REGION Network 3: Convoyeur 02
   RUNG wire#powerrail
      #Convoyeur_Hippodrome_2(x_Marche_auto := wire#w1, x_Arret_auto := wire#w2, x_Defaut_externe := "Bits_Globaux".x_Defaut_bloquant, x_enService := "Bits_Globaux".x_En_service, x_Marche_manu := "Tch_HMI".Tch_Manu[50], x_Arret_Manu := "Tch_HMI".Tch_Manu[51], x_Retour_defaut_thermique := "I_Def_Thermique_CV02_hyppo", DB_Convoyeur_DATA := "DB_Convoyeurs_Hipp".Convoyeur[2], Defaut =>)
   END_RUNG
   RUNG wire#powerrail
      Contact( "Bits_Globaux".x_En_cycle_auto )
   END_RUNG wire#w1
   RUNG wire#powerrail
      Contact( "Bits_Globaux".x_Demo_Hippo_en_cours )
   END_RUNG wire#w1
   RUNG wire#powerrail
      Contact( "Tch_HMI".Tch_Acy )
   END_RUNG wire#w2
   RUNG wire#powerrail
      Contact( #x_All_stations_empty )
   END_RUNG wire#w2
   // the same network as SCL:
   #Convoyeur_Hippodrome_2(x_Defaut_externe := "Bits_Globaux".x_Defaut_bloquant,   // "Convoyeur_Hippodrome"
                           x_enService := "Bits_Globaux".x_En_service,
                           x_Marche_auto := "Bits_Globaux".x_En_cycle_auto OR "Bits_Globaux".x_Demo_Hippo_en_cours,
                           x_Marche_manu := "Tch_HMI".Tch_Manu[50],
                           x_Arret_auto := "Tch_HMI".Tch_Acy OR #x_All_stations_empty,
                           x_Arret_Manu := "Tch_HMI".Tch_Manu[51],
                           x_Retour_defaut_thermique := "I_Def_Thermique_CV02_hyppo",
                           DB_Convoyeur_DATA := "DB_Convoyeurs_Hipp".Convoyeur[2]);
END_REGION

REGION Network 4: Convoyeur 03
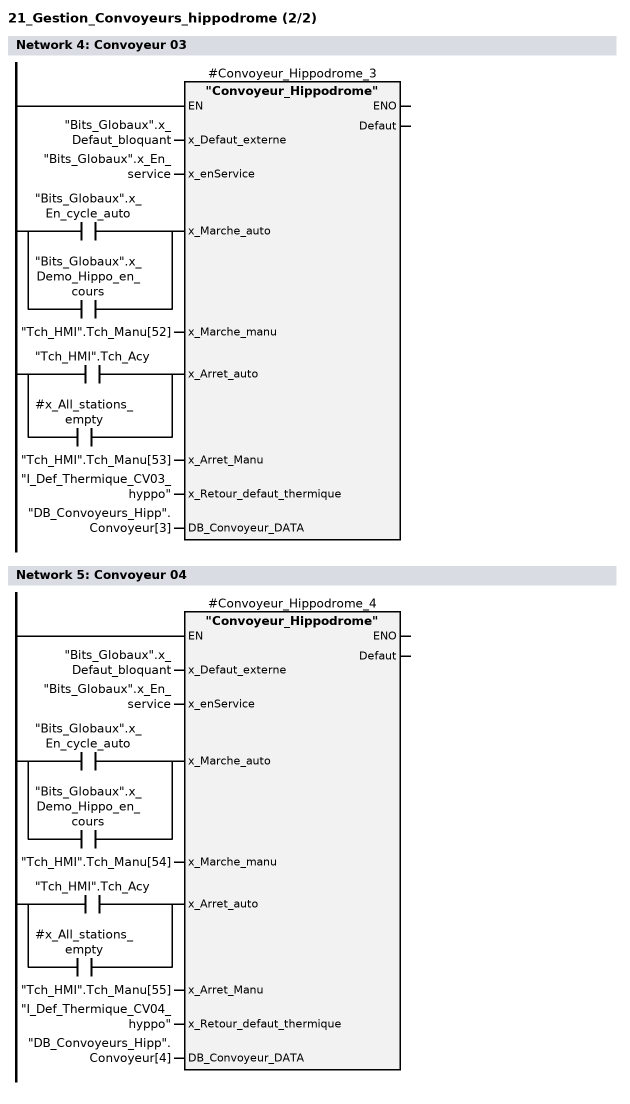
   RUNG wire#powerrail
      #Convoyeur_Hippodrome_3(x_Marche_auto := wire#w1, x_Arret_auto := wire#w2, x_Defaut_externe := "Bits_Globaux".x_Defaut_bloquant, x_enService := "Bits_Globaux".x_En_service, x_Marche_manu := "Tch_HMI".Tch_Manu[52], x_Arret_Manu := "Tch_HMI".Tch_Manu[53], x_Retour_defaut_thermique := "I_Def_Thermique_CV03_hyppo", DB_Convoyeur_DATA := "DB_Convoyeurs_Hipp".Convoyeur[3], Defaut =>)
   END_RUNG
   RUNG wire#powerrail
      Contact( "Bits_Globaux".x_En_cycle_auto )
   END_RUNG wire#w1
   RUNG wire#powerrail
      Contact( "Bits_Globaux".x_Demo_Hippo_en_cours )
   END_RUNG wire#w1
   RUNG wire#powerrail
      Contact( "Tch_HMI".Tch_Acy )
   END_RUNG wire#w2
   RUNG wire#powerrail
      Contact( #x_All_stations_empty )
   END_RUNG wire#w2
   // the same network as SCL:
   #Convoyeur_Hippodrome_3(x_Defaut_externe := "Bits_Globaux".x_Defaut_bloquant,   // "Convoyeur_Hippodrome"
                           x_enService := "Bits_Globaux".x_En_service,
                           x_Marche_auto := "Bits_Globaux".x_En_cycle_auto OR "Bits_Globaux".x_Demo_Hippo_en_cours,
                           x_Marche_manu := "Tch_HMI".Tch_Manu[52],
                           x_Arret_auto := "Tch_HMI".Tch_Acy OR #x_All_stations_empty,
                           x_Arret_Manu := "Tch_HMI".Tch_Manu[53],
                           x_Retour_defaut_thermique := "I_Def_Thermique_CV03_hyppo",
                           DB_Convoyeur_DATA := "DB_Convoyeurs_Hipp".Convoyeur[3]);
END_REGION

REGION Network 5: Convoyeur 04
   RUNG wire#powerrail
      #Convoyeur_Hippodrome_4(x_Marche_auto := wire#w1, x_Arret_auto := wire#w2, x_Defaut_externe := "Bits_Globaux".x_Defaut_bloquant, x_enService := "Bits_Globaux".x_En_service, x_Marche_manu := "Tch_HMI".Tch_Manu[54], x_Arret_Manu := "Tch_HMI".Tch_Manu[55], x_Retour_defaut_thermique := "I_Def_Thermique_CV04_hyppo", DB_Convoyeur_DATA := "DB_Convoyeurs_Hipp".Convoyeur[4], Defaut =>)
   END_RUNG
   RUNG wire#powerrail
      Contact( "Bits_Globaux".x_En_cycle_auto )
   END_RUNG wire#w1
   RUNG wire#powerrail
      Contact( "Bits_Globaux".x_Demo_Hippo_en_cours )
   END_RUNG wire#w1
   RUNG wire#powerrail
      Contact( "Tch_HMI".Tch_Acy )
   END_RUNG wire#w2
   RUNG wire#powerrail
      Contact( #x_All_stations_empty )
   END_RUNG wire#w2
   // the same network as SCL:
   #Convoyeur_Hippodrome_4(x_Defaut_externe := "Bits_Globaux".x_Defaut_bloquant,   // "Convoyeur_Hippodrome"
                           x_enService := "Bits_Globaux".x_En_service,
                           x_Marche_auto := "Bits_Globaux".x_En_cycle_auto OR "Bits_Globaux".x_Demo_Hippo_en_cours,
                           x_Marche_manu := "Tch_HMI".Tch_Manu[54],
                           x_Arret_auto := "Tch_HMI".Tch_Acy OR #x_All_stations_empty,
                           x_Arret_Manu := "Tch_HMI".Tch_Manu[55],
                           x_Retour_defaut_thermique := "I_Def_Thermique_CV04_hyppo",
                           DB_Convoyeur_DATA := "DB_Convoyeurs_Hipp".Convoyeur[4]);
END_REGION
END_FUNCTION_BLOCK

// folder: 2-Hippodrome/Stations de travail

FUNCTION_BLOCK "22-Gestion_stations"   // FB10, LAD
{ S7_Optimized_Access := 'TRUE' }
VERSION : 0.1
   VAR
      Station_de_travail_1 : "Station_de_travail";
      Station_de_travail_2 : "Station_de_travail";
      Station_de_travail_3 : "Station_de_travail";
      Station_de_travail_4 : "Station_de_travail";
      Station_de_travail_5 : "Station_de_travail";
      Station_de_travail_6 : "Station_de_travail";
      Station_de_travail_7 : "Station_de_travail";
      x_WorkDone_mode_demo : Bool;
      Front_montant_Demo_1 : Bool;
      Timer_front_montant : TP_TIME;
      x_All_stations_empty : Bool;
   END_VAR
   VAR_TEMP   // added for the SCL form of the ladder/FBD networks
      _w1 : Bool;
   END_VAR
BEGIN

REGION Network 1: Gestion palettes si toutes les palettes son vides
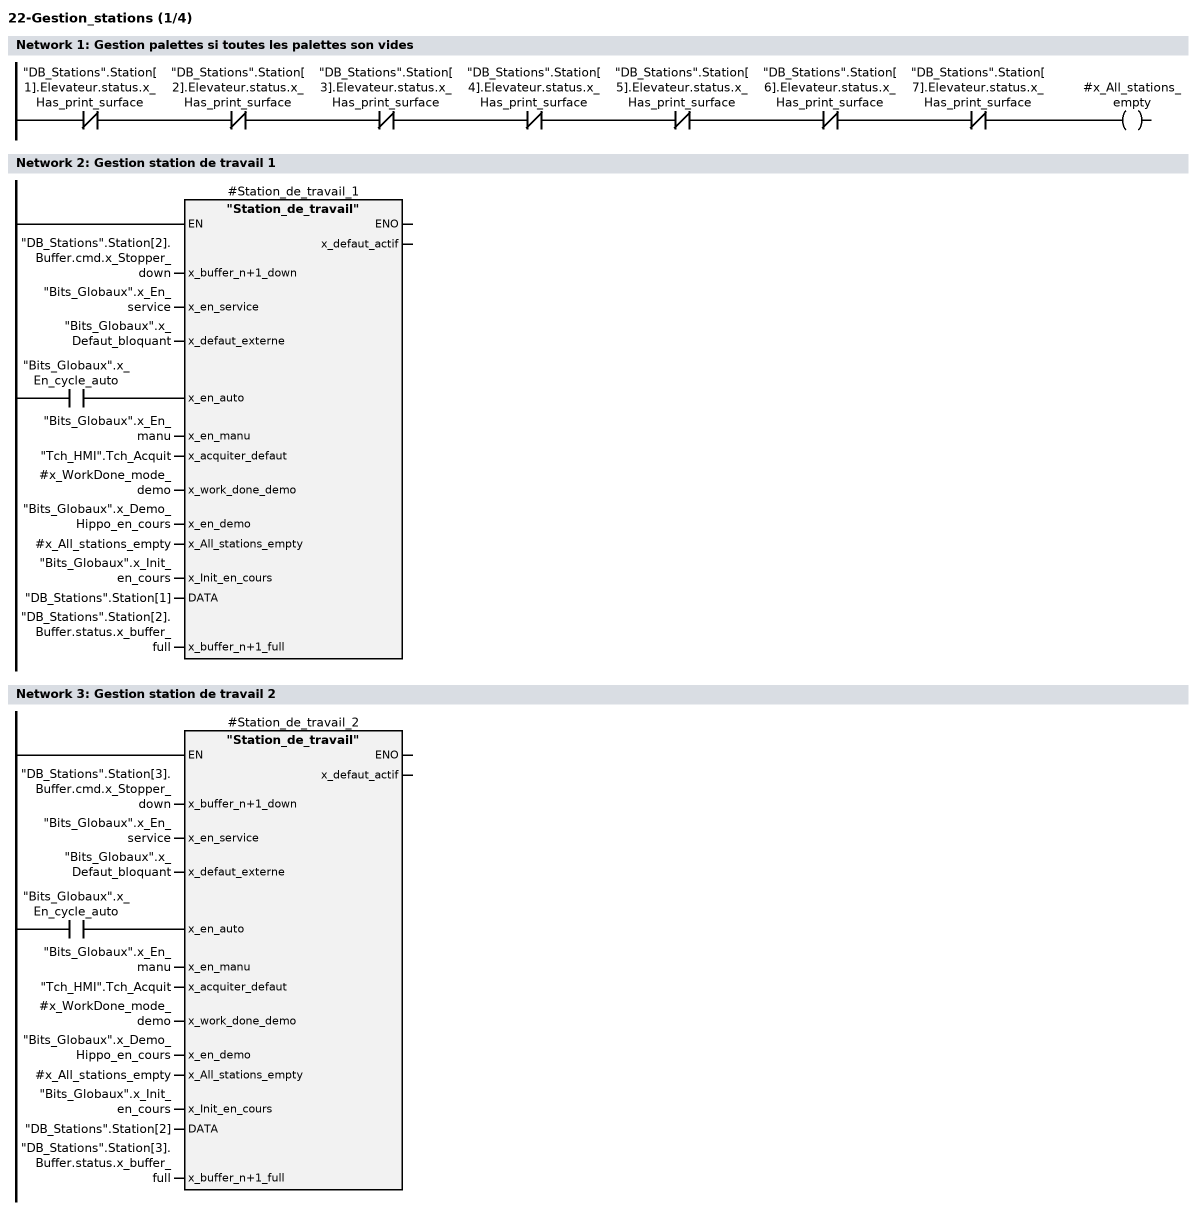
   RUNG wire#powerrail
      I_Contact( "DB_Stations".Station[1].Elevateur.status.x_Has_print_surface )
      I_Contact( "DB_Stations".Station[2].Elevateur.status.x_Has_print_surface )
      I_Contact( "DB_Stations".Station[3].Elevateur.status.x_Has_print_surface )
      I_Contact( "DB_Stations".Station[4].Elevateur.status.x_Has_print_surface )
      I_Contact( "DB_Stations".Station[5].Elevateur.status.x_Has_print_surface )
      I_Contact( "DB_Stations".Station[6].Elevateur.status.x_Has_print_surface )
      I_Contact( "DB_Stations".Station[7].Elevateur.status.x_Has_print_surface )
      Coil( #x_All_stations_empty )
   END_RUNG
   // the same network as SCL:
   #x_All_stations_empty := NOT "DB_Stations".Station[1].Elevateur.status.x_Has_print_surface AND NOT "DB_Stations".Station[2].Elevateur.status.x_Has_print_surface AND NOT "DB_Stations".Station[3].Elevateur.status.x_Has_print_surface AND NOT "DB_Stations".Station[4].Elevateur.status.x_Has_print_surface AND NOT "DB_Stations".Station[5].Elevateur.status.x_Has_print_surface AND NOT "DB_Stations".Station[6].Elevateur.status.x_Has_print_surface AND NOT "DB_Stations".Station[7].Elevateur.status.x_Has_print_surface;
END_REGION

REGION Network 2: Gestion station de travail 1
   RUNG wire#powerrail
      #Station_de_travail_1(x_en_auto := wire#w1, "x_buffer_n+1_down" := "DB_Stations".Station[2].Buffer.cmd.x_Stopper_down, x_en_service := "Bits_Globaux".x_En_service, x_defaut_externe := "Bits_Globaux".x_Defaut_bloquant, x_en_manu := "Bits_Globaux".x_En_manu, x_acquiter_defaut := "Tch_HMI".Tch_Acquit, x_work_done_demo := #x_WorkDone_mode_demo, x_en_demo := "Bits_Globaux".x_Demo_Hippo_en_cours, x_All_stations_empty := #x_All_stations_empty, x_Init_en_cours := "Bits_Globaux".x_Init_en_cours, DATA := "DB_Stations".Station[1], "x_buffer_n+1_full" := "DB_Stations".Station[2].Buffer.status.x_buffer_full, x_defaut_actif =>)
   END_RUNG
   RUNG wire#powerrail
      Contact( "Bits_Globaux".x_En_cycle_auto )
   END_RUNG wire#w1
   // the same network as SCL:
   #Station_de_travail_1("x_buffer_n+1_down" := "DB_Stations".Station[2].Buffer.cmd.x_Stopper_down,   // "Station_de_travail"
                         x_en_service := "Bits_Globaux".x_En_service,
                         x_defaut_externe := "Bits_Globaux".x_Defaut_bloquant,
                         x_en_auto := "Bits_Globaux".x_En_cycle_auto,
                         x_en_manu := "Bits_Globaux".x_En_manu,
                         x_acquiter_defaut := "Tch_HMI".Tch_Acquit,
                         x_work_done_demo := #x_WorkDone_mode_demo,
                         x_en_demo := "Bits_Globaux".x_Demo_Hippo_en_cours,
                         x_All_stations_empty := #x_All_stations_empty,
                         x_Init_en_cours := "Bits_Globaux".x_Init_en_cours,
                         DATA := "DB_Stations".Station[1],
                         "x_buffer_n+1_full" := "DB_Stations".Station[2].Buffer.status.x_buffer_full);
END_REGION

REGION Network 3: Gestion station de travail 2
   RUNG wire#powerrail
      #Station_de_travail_2(x_en_auto := wire#w1, "x_buffer_n+1_down" := "DB_Stations".Station[3].Buffer.cmd.x_Stopper_down, x_en_service := "Bits_Globaux".x_En_service, x_defaut_externe := "Bits_Globaux".x_Defaut_bloquant, x_en_manu := "Bits_Globaux".x_En_manu, x_acquiter_defaut := "Tch_HMI".Tch_Acquit, x_work_done_demo := #x_WorkDone_mode_demo, x_en_demo := "Bits_Globaux".x_Demo_Hippo_en_cours, x_All_stations_empty := #x_All_stations_empty, x_Init_en_cours := "Bits_Globaux".x_Init_en_cours, DATA := "DB_Stations".Station[2], "x_buffer_n+1_full" := "DB_Stations".Station[3].Buffer.status.x_buffer_full, x_defaut_actif =>)
   END_RUNG
   RUNG wire#powerrail
      Contact( "Bits_Globaux".x_En_cycle_auto )
   END_RUNG wire#w1
   // the same network as SCL:
   #Station_de_travail_2("x_buffer_n+1_down" := "DB_Stations".Station[3].Buffer.cmd.x_Stopper_down,   // "Station_de_travail"
                         x_en_service := "Bits_Globaux".x_En_service,
                         x_defaut_externe := "Bits_Globaux".x_Defaut_bloquant,
                         x_en_auto := "Bits_Globaux".x_En_cycle_auto,
                         x_en_manu := "Bits_Globaux".x_En_manu,
                         x_acquiter_defaut := "Tch_HMI".Tch_Acquit,
                         x_work_done_demo := #x_WorkDone_mode_demo,
                         x_en_demo := "Bits_Globaux".x_Demo_Hippo_en_cours,
                         x_All_stations_empty := #x_All_stations_empty,
                         x_Init_en_cours := "Bits_Globaux".x_Init_en_cours,
                         DATA := "DB_Stations".Station[2],
                         "x_buffer_n+1_full" := "DB_Stations".Station[3].Buffer.status.x_buffer_full);
END_REGION

REGION Network 4: Gestion station de travail 3
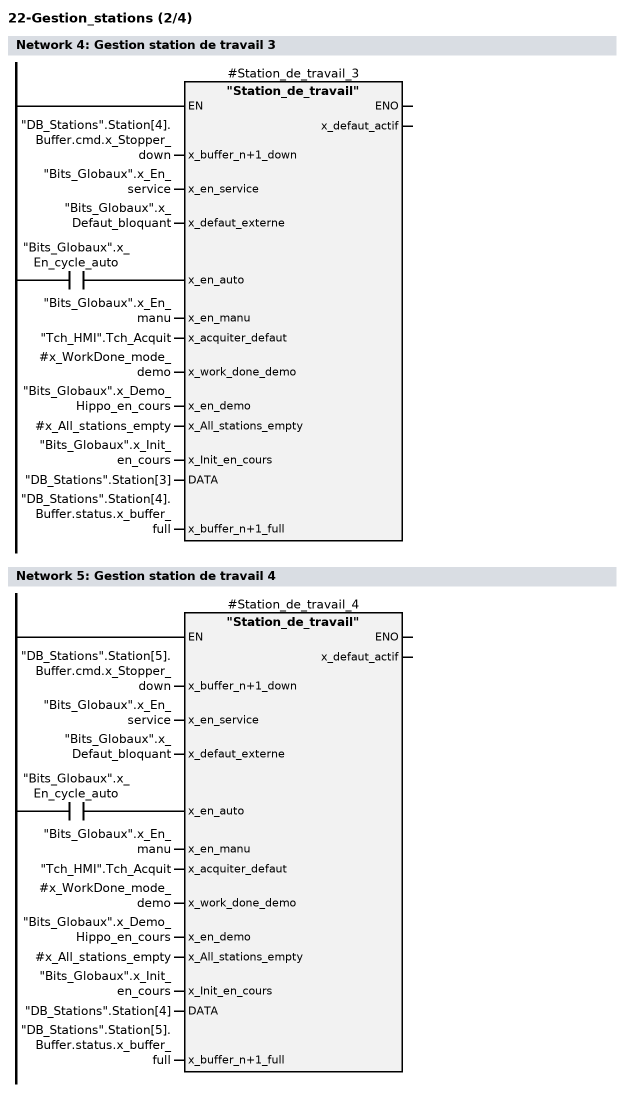
   RUNG wire#powerrail
      #Station_de_travail_3(x_en_auto := wire#w1, "x_buffer_n+1_down" := "DB_Stations".Station[4].Buffer.cmd.x_Stopper_down, x_en_service := "Bits_Globaux".x_En_service, x_defaut_externe := "Bits_Globaux".x_Defaut_bloquant, x_en_manu := "Bits_Globaux".x_En_manu, x_acquiter_defaut := "Tch_HMI".Tch_Acquit, x_work_done_demo := #x_WorkDone_mode_demo, x_en_demo := "Bits_Globaux".x_Demo_Hippo_en_cours, x_All_stations_empty := #x_All_stations_empty, x_Init_en_cours := "Bits_Globaux".x_Init_en_cours, DATA := "DB_Stations".Station[3], "x_buffer_n+1_full" := "DB_Stations".Station[4].Buffer.status.x_buffer_full, x_defaut_actif =>)
   END_RUNG
   RUNG wire#powerrail
      Contact( "Bits_Globaux".x_En_cycle_auto )
   END_RUNG wire#w1
   // the same network as SCL:
   #Station_de_travail_3("x_buffer_n+1_down" := "DB_Stations".Station[4].Buffer.cmd.x_Stopper_down,   // "Station_de_travail"
                         x_en_service := "Bits_Globaux".x_En_service,
                         x_defaut_externe := "Bits_Globaux".x_Defaut_bloquant,
                         x_en_auto := "Bits_Globaux".x_En_cycle_auto,
                         x_en_manu := "Bits_Globaux".x_En_manu,
                         x_acquiter_defaut := "Tch_HMI".Tch_Acquit,
                         x_work_done_demo := #x_WorkDone_mode_demo,
                         x_en_demo := "Bits_Globaux".x_Demo_Hippo_en_cours,
                         x_All_stations_empty := #x_All_stations_empty,
                         x_Init_en_cours := "Bits_Globaux".x_Init_en_cours,
                         DATA := "DB_Stations".Station[3],
                         "x_buffer_n+1_full" := "DB_Stations".Station[4].Buffer.status.x_buffer_full);
END_REGION

REGION Network 5: Gestion station de travail 4
   RUNG wire#powerrail
      #Station_de_travail_4(x_en_auto := wire#w1, "x_buffer_n+1_down" := "DB_Stations".Station[5].Buffer.cmd.x_Stopper_down, x_en_service := "Bits_Globaux".x_En_service, x_defaut_externe := "Bits_Globaux".x_Defaut_bloquant, x_en_manu := "Bits_Globaux".x_En_manu, x_acquiter_defaut := "Tch_HMI".Tch_Acquit, x_work_done_demo := #x_WorkDone_mode_demo, x_en_demo := "Bits_Globaux".x_Demo_Hippo_en_cours, x_All_stations_empty := #x_All_stations_empty, x_Init_en_cours := "Bits_Globaux".x_Init_en_cours, DATA := "DB_Stations".Station[4], "x_buffer_n+1_full" := "DB_Stations".Station[5].Buffer.status.x_buffer_full, x_defaut_actif =>)
   END_RUNG
   RUNG wire#powerrail
      Contact( "Bits_Globaux".x_En_cycle_auto )
   END_RUNG wire#w1
   // the same network as SCL:
   #Station_de_travail_4("x_buffer_n+1_down" := "DB_Stations".Station[5].Buffer.cmd.x_Stopper_down,   // "Station_de_travail"
                         x_en_service := "Bits_Globaux".x_En_service,
                         x_defaut_externe := "Bits_Globaux".x_Defaut_bloquant,
                         x_en_auto := "Bits_Globaux".x_En_cycle_auto,
                         x_en_manu := "Bits_Globaux".x_En_manu,
                         x_acquiter_defaut := "Tch_HMI".Tch_Acquit,
                         x_work_done_demo := #x_WorkDone_mode_demo,
                         x_en_demo := "Bits_Globaux".x_Demo_Hippo_en_cours,
                         x_All_stations_empty := #x_All_stations_empty,
                         x_Init_en_cours := "Bits_Globaux".x_Init_en_cours,
                         DATA := "DB_Stations".Station[4],
                         "x_buffer_n+1_full" := "DB_Stations".Station[5].Buffer.status.x_buffer_full);
END_REGION

REGION Network 6: Gestion station de travail 5
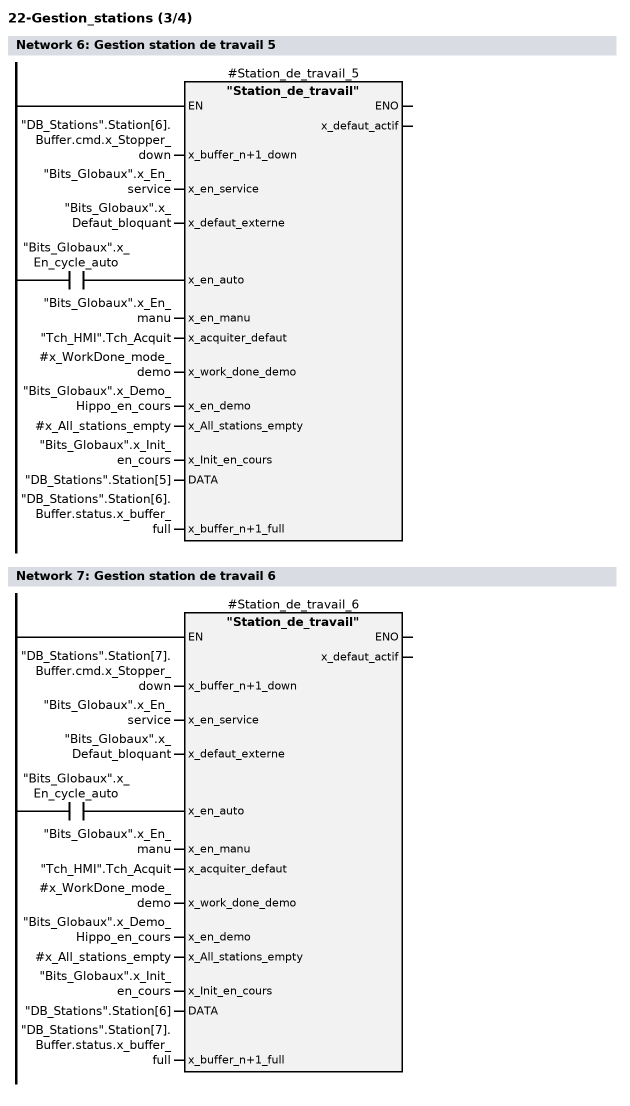
   RUNG wire#powerrail
      #Station_de_travail_5(x_en_auto := wire#w1, "x_buffer_n+1_down" := "DB_Stations".Station[6].Buffer.cmd.x_Stopper_down, x_en_service := "Bits_Globaux".x_En_service, x_defaut_externe := "Bits_Globaux".x_Defaut_bloquant, x_en_manu := "Bits_Globaux".x_En_manu, x_acquiter_defaut := "Tch_HMI".Tch_Acquit, x_work_done_demo := #x_WorkDone_mode_demo, x_en_demo := "Bits_Globaux".x_Demo_Hippo_en_cours, x_All_stations_empty := #x_All_stations_empty, x_Init_en_cours := "Bits_Globaux".x_Init_en_cours, DATA := "DB_Stations".Station[5], "x_buffer_n+1_full" := "DB_Stations".Station[6].Buffer.status.x_buffer_full, x_defaut_actif =>)
   END_RUNG
   RUNG wire#powerrail
      Contact( "Bits_Globaux".x_En_cycle_auto )
   END_RUNG wire#w1
   // the same network as SCL:
   #Station_de_travail_5("x_buffer_n+1_down" := "DB_Stations".Station[6].Buffer.cmd.x_Stopper_down,   // "Station_de_travail"
                         x_en_service := "Bits_Globaux".x_En_service,
                         x_defaut_externe := "Bits_Globaux".x_Defaut_bloquant,
                         x_en_auto := "Bits_Globaux".x_En_cycle_auto,
                         x_en_manu := "Bits_Globaux".x_En_manu,
                         x_acquiter_defaut := "Tch_HMI".Tch_Acquit,
                         x_work_done_demo := #x_WorkDone_mode_demo,
                         x_en_demo := "Bits_Globaux".x_Demo_Hippo_en_cours,
                         x_All_stations_empty := #x_All_stations_empty,
                         x_Init_en_cours := "Bits_Globaux".x_Init_en_cours,
                         DATA := "DB_Stations".Station[5],
                         "x_buffer_n+1_full" := "DB_Stations".Station[6].Buffer.status.x_buffer_full);
END_REGION

REGION Network 7: Gestion station de travail 6
   RUNG wire#powerrail
      #Station_de_travail_6(x_en_auto := wire#w1, "x_buffer_n+1_down" := "DB_Stations".Station[7].Buffer.cmd.x_Stopper_down, x_en_service := "Bits_Globaux".x_En_service, x_defaut_externe := "Bits_Globaux".x_Defaut_bloquant, x_en_manu := "Bits_Globaux".x_En_manu, x_acquiter_defaut := "Tch_HMI".Tch_Acquit, x_work_done_demo := #x_WorkDone_mode_demo, x_en_demo := "Bits_Globaux".x_Demo_Hippo_en_cours, x_All_stations_empty := #x_All_stations_empty, x_Init_en_cours := "Bits_Globaux".x_Init_en_cours, DATA := "DB_Stations".Station[6], "x_buffer_n+1_full" := "DB_Stations".Station[7].Buffer.status.x_buffer_full, x_defaut_actif =>)
   END_RUNG
   RUNG wire#powerrail
      Contact( "Bits_Globaux".x_En_cycle_auto )
   END_RUNG wire#w1
   // the same network as SCL:
   #Station_de_travail_6("x_buffer_n+1_down" := "DB_Stations".Station[7].Buffer.cmd.x_Stopper_down,   // "Station_de_travail"
                         x_en_service := "Bits_Globaux".x_En_service,
                         x_defaut_externe := "Bits_Globaux".x_Defaut_bloquant,
                         x_en_auto := "Bits_Globaux".x_En_cycle_auto,
                         x_en_manu := "Bits_Globaux".x_En_manu,
                         x_acquiter_defaut := "Tch_HMI".Tch_Acquit,
                         x_work_done_demo := #x_WorkDone_mode_demo,
                         x_en_demo := "Bits_Globaux".x_Demo_Hippo_en_cours,
                         x_All_stations_empty := #x_All_stations_empty,
                         x_Init_en_cours := "Bits_Globaux".x_Init_en_cours,
                         DATA := "DB_Stations".Station[6],
                         "x_buffer_n+1_full" := "DB_Stations".Station[7].Buffer.status.x_buffer_full);
END_REGION

REGION Network 8: Gestion station de travail 7
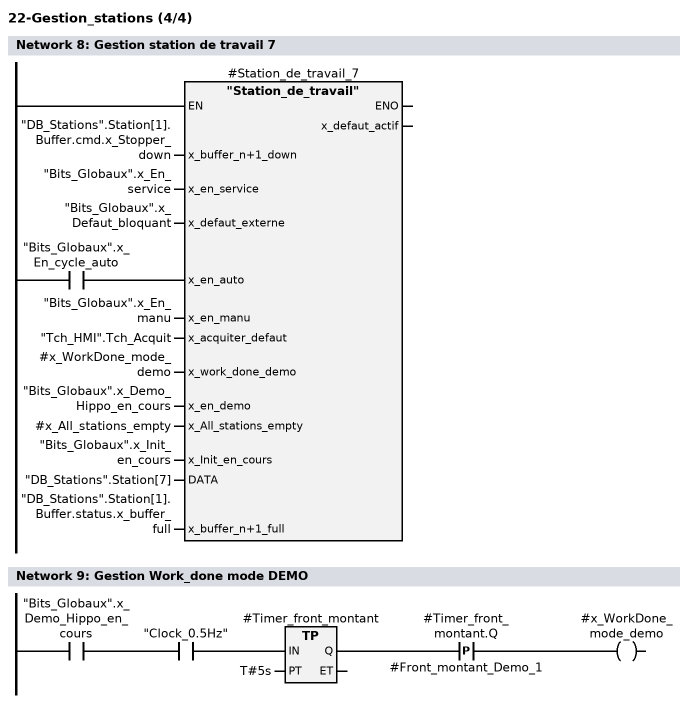
   RUNG wire#powerrail
      #Station_de_travail_7(x_en_auto := wire#w1, "x_buffer_n+1_down" := "DB_Stations".Station[1].Buffer.cmd.x_Stopper_down, x_en_service := "Bits_Globaux".x_En_service, x_defaut_externe := "Bits_Globaux".x_Defaut_bloquant, x_en_manu := "Bits_Globaux".x_En_manu, x_acquiter_defaut := "Tch_HMI".Tch_Acquit, x_work_done_demo := #x_WorkDone_mode_demo, x_en_demo := "Bits_Globaux".x_Demo_Hippo_en_cours, x_All_stations_empty := #x_All_stations_empty, x_Init_en_cours := "Bits_Globaux".x_Init_en_cours, DATA := "DB_Stations".Station[7], "x_buffer_n+1_full" := "DB_Stations".Station[1].Buffer.status.x_buffer_full, x_defaut_actif =>)
   END_RUNG
   RUNG wire#powerrail
      Contact( "Bits_Globaux".x_En_cycle_auto )
   END_RUNG wire#w1
   // the same network as SCL:
   #Station_de_travail_7("x_buffer_n+1_down" := "DB_Stations".Station[1].Buffer.cmd.x_Stopper_down,   // "Station_de_travail"
                         x_en_service := "Bits_Globaux".x_En_service,
                         x_defaut_externe := "Bits_Globaux".x_Defaut_bloquant,
                         x_en_auto := "Bits_Globaux".x_En_cycle_auto,
                         x_en_manu := "Bits_Globaux".x_En_manu,
                         x_acquiter_defaut := "Tch_HMI".Tch_Acquit,
                         x_work_done_demo := #x_WorkDone_mode_demo,
                         x_en_demo := "Bits_Globaux".x_Demo_Hippo_en_cours,
                         x_All_stations_empty := #x_All_stations_empty,
                         x_Init_en_cours := "Bits_Globaux".x_Init_en_cours,
                         DATA := "DB_Stations".Station[7],
                         "x_buffer_n+1_full" := "DB_Stations".Station[1].Buffer.status.x_buffer_full);
END_REGION

REGION Network 9: Gestion Work_done mode DEMO
   #Timer_front_montant(IN := "Bits_Globaux".x_Demo_Hippo_en_cours AND "Clock_0.5Hz", PT := T#5s);   // TP
   #_w1 := #Timer_front_montant.Q AND #Timer_front_montant.Q AND NOT #Front_montant_Demo_1;   // rising edge of #Timer_front_montant.Q
   #Front_montant_Demo_1 := #Timer_front_montant.Q;
   #x_WorkDone_mode_demo := #_w1;
END_REGION
END_FUNCTION_BLOCK

FUNCTION_BLOCK "Station_de_travail"   // FB11, LAD
TITLE = Controle Station de travail
{ S7_Optimized_Access := 'TRUE' }
VERSION : 0.1
   VAR_INPUT
      "x_buffer_n+1_down" : Bool;
      x_en_service : Bool;
      x_defaut_externe : Bool;
      x_en_auto : Bool;
      x_en_manu : Bool;
      x_acquiter_defaut : Bool;
      x_work_done_demo : Bool;
      x_en_demo : Bool;
      x_All_stations_empty : Bool;
      x_Init_en_cours : Bool;
   END_VAR
   VAR_OUTPUT
      x_defaut_actif : Bool;
   END_VAR
   VAR_IN_OUT
      DATA : "Station_Hipp";
      "x_buffer_n+1_full" : Bool;
   END_VAR
   VAR
      Front_descendant_presence_elevateur : Bool;
      Front_descendant_presence_buffer : Bool;
   END_VAR
   VAR RETAIN
      Instance_Compteur_sortie_EL : CTU_INT;
   END_VAR
   VAR
      IEC_Timer_Delai_remontee_butee_el : TON_TIME;
      IEC_Timer_0_Instance_1 : TON_TIME;
      IEC_Timer_Discordance_descente : TON_TIME;
      IEC_Timer_Discordance_montee : TON_TIME;
      Front_descendant_butee_elevateur : Bool;
      Front_descendant_descente_EL : Bool;
      Front_descendant_descente_EL_2 : Bool;
      Front_montant_etat_free : Bool;
      Front_descendant_timer_butee_El : Bool;
      IEC_Timer_0_Instance : TP_TIME;
      IEC_Timer_0_Instance_2 : TON_TIME;
      Timer_ByPassDemo_ElevatorDown : TON_TIME;
   END_VAR
   VAR_TEMP   // added for the SCL form of the ladder/FBD networks
      _w1 : Bool;
      _w2 : Bool;
   END_VAR
BEGIN

REGION Network 1: Gestion butee buffer
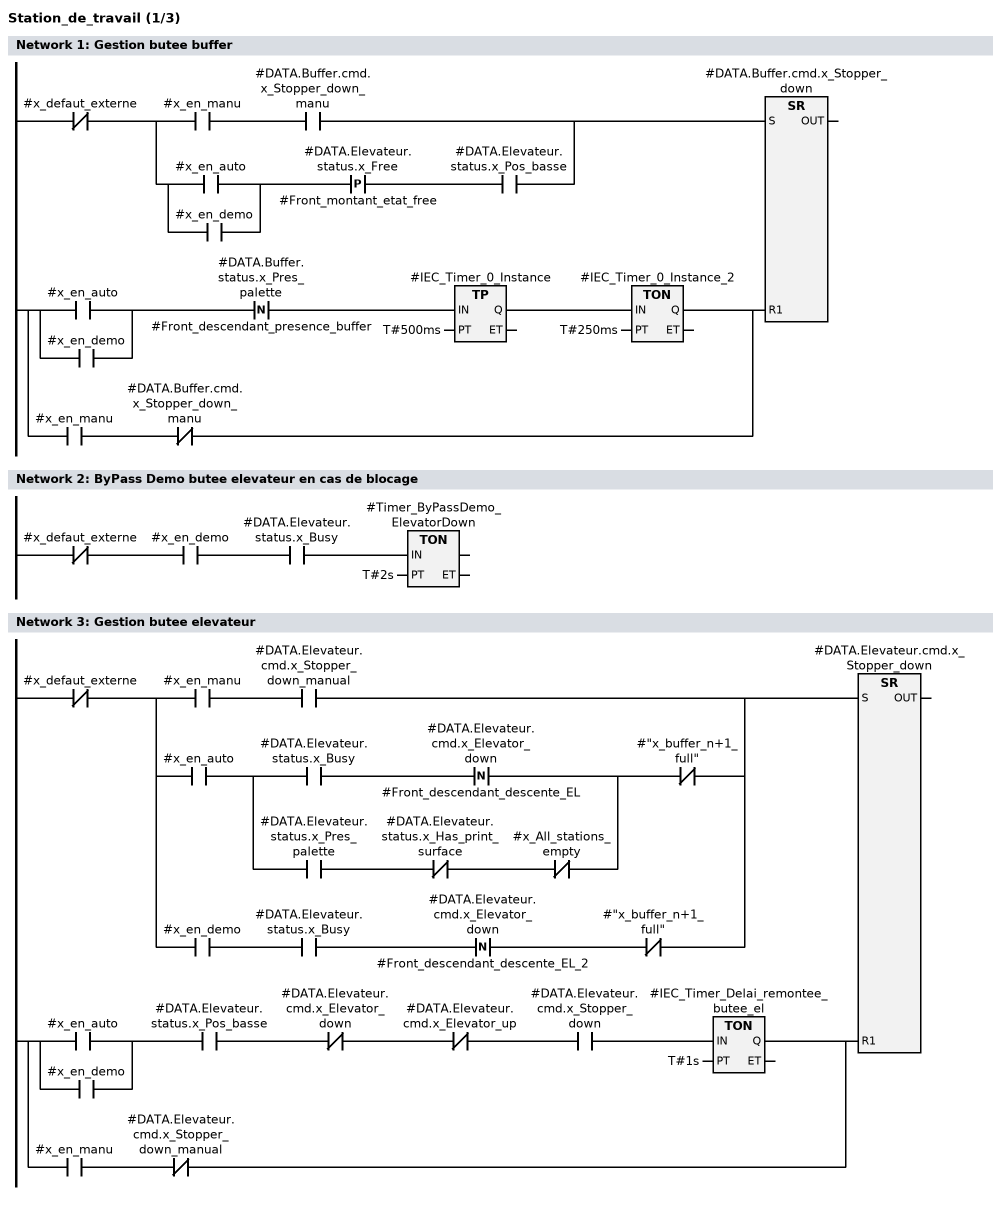
   #_w1 := NOT #x_defaut_externe AND (#x_en_auto OR #x_en_demo) AND #DATA.Elevateur.status.x_Free AND NOT #Front_montant_etat_free;   // rising edge of #DATA.Elevateur.status.x_Free
   #Front_montant_etat_free := #DATA.Elevateur.status.x_Free;
   #_w2 := (#x_en_auto OR #x_en_demo) AND NOT #DATA.Buffer.status.x_Pres_palette AND #Front_descendant_presence_buffer;   // falling edge of #DATA.Buffer.status.x_Pres_palette
   #Front_descendant_presence_buffer := #DATA.Buffer.status.x_Pres_palette;
   #IEC_Timer_0_Instance(IN := #_w2, PT := T#500ms);   // TP
   #IEC_Timer_0_Instance_2(IN := #IEC_Timer_0_Instance.Q, PT := T#250ms);   // TON
   IF (NOT #x_defaut_externe AND #x_en_manu AND #DATA.Buffer.cmd.x_Stopper_down_manu) OR (#_w1 AND #DATA.Elevateur.status.x_Pos_basse) THEN
       #DATA.Buffer.cmd.x_Stopper_down := TRUE;   // SR flip-flop
   END_IF;
   IF #IEC_Timer_0_Instance_2.Q OR (#x_en_manu AND NOT #DATA.Buffer.cmd.x_Stopper_down_manu) THEN
       #DATA.Buffer.cmd.x_Stopper_down := FALSE;
   END_IF;
END_REGION

REGION Network 2: ByPass Demo butee elevateur en cas de blocage
   #Timer_ByPassDemo_ElevatorDown(IN := NOT #x_defaut_externe AND #x_en_demo AND #DATA.Elevateur.status.x_Busy,   // TON
                           PT := T#2s);
END_REGION

REGION Network 3: Gestion butee elevateur
   #_w1 := NOT #x_defaut_externe AND #x_en_auto AND #DATA.Elevateur.status.x_Busy AND NOT #DATA.Elevateur.cmd.x_Elevator_down AND #Front_descendant_descente_EL;   // falling edge of #DATA.Elevateur.cmd.x_Elevator_down
   #Front_descendant_descente_EL := #DATA.Elevateur.cmd.x_Elevator_down;
   #_w2 := NOT #x_defaut_externe AND #x_en_demo AND #DATA.Elevateur.status.x_Busy AND NOT #DATA.Elevateur.cmd.x_Elevator_down AND #Front_descendant_descente_EL_2;   // falling edge of #DATA.Elevateur.cmd.x_Elevator_down
   #Front_descendant_descente_EL_2 := #DATA.Elevateur.cmd.x_Elevator_down;
   #IEC_Timer_Delai_remontee_butee_el(IN := (#x_en_auto OR #x_en_demo) AND #DATA.Elevateur.status.x_Pos_basse AND NOT #DATA.Elevateur.cmd.x_Elevator_down AND NOT #DATA.Elevateur.cmd.x_Elevator_up AND #DATA.Elevateur.cmd.x_Stopper_down,   // TON
                           PT := T#1s);
   IF (NOT #x_defaut_externe AND #x_en_manu AND #DATA.Elevateur.cmd.x_Stopper_down_manual) OR ((#_w1 OR (NOT #x_defaut_externe AND #x_en_auto AND #DATA.Elevateur.status.x_Pres_palette AND NOT #DATA.Elevateur.status.x_Has_print_surface AND NOT #x_All_stations_empty)) AND NOT #"x_buffer_n+1_full") OR (#_w2 AND NOT #"x_buffer_n+1_full") THEN
       #DATA.Elevateur.cmd.x_Stopper_down := TRUE;   // SR flip-flop
   END_IF;
   IF #IEC_Timer_Delai_remontee_butee_el.Q OR (#x_en_manu AND NOT #DATA.Elevateur.cmd.x_Stopper_down_manual) THEN
       #DATA.Elevateur.cmd.x_Stopper_down := FALSE;
   END_IF;
END_REGION

REGION Network 4: Gestion compteur palettes sur buffer n+1
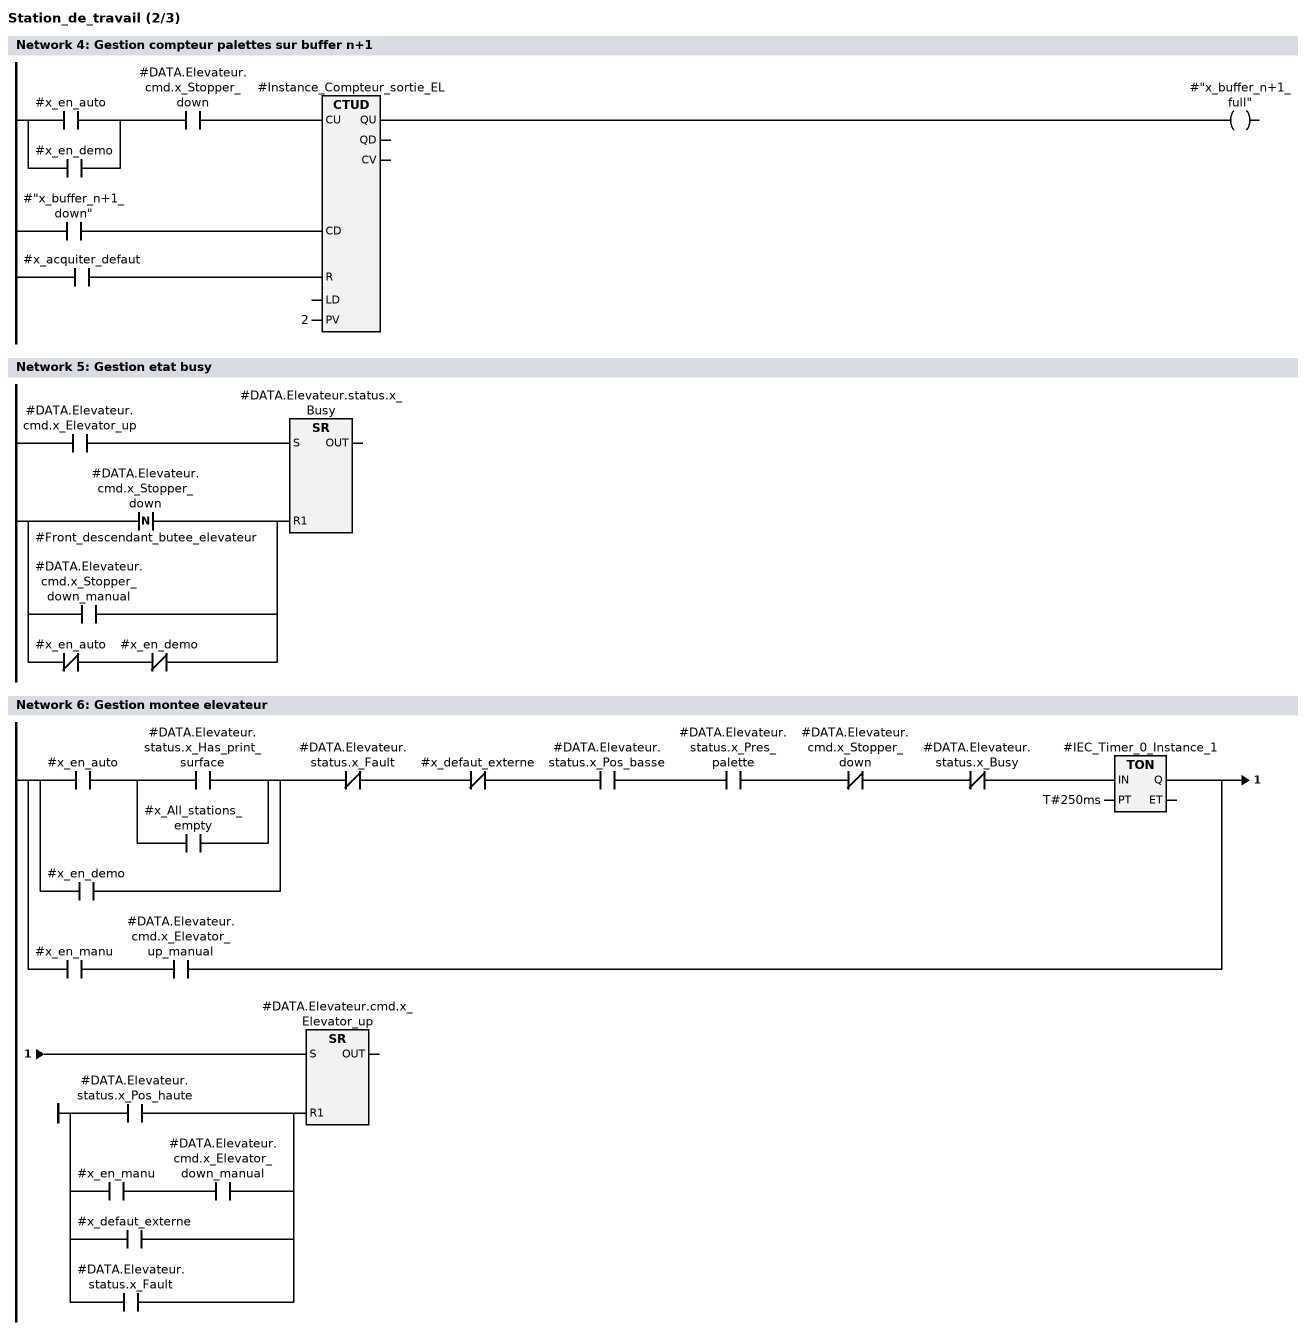
   #Instance_Compteur_sortie_EL(CU := (#x_en_auto OR #x_en_demo) AND #DATA.Elevateur.cmd.x_Stopper_down,   // CTUD
                           CD := #"x_buffer_n+1_down",
                           R := #x_acquiter_defaut,
                           PV := 2);
   #"x_buffer_n+1_full" := #Instance_Compteur_sortie_EL.QU;
END_REGION

REGION Network 5: Gestion etat busy
   RUNG wire#powerrail
      Contact( #DATA.Elevateur.cmd.x_Elevator_up )
      S_SR(operand := #DATA.Elevateur.status.x_Busy, r1 := wire#w1)
   END_RUNG
   RUNG wire#powerrail
      N_Contact(operand := #DATA.Elevateur.cmd.x_Stopper_down, bit := #Front_descendant_butee_elevateur)
   END_RUNG wire#w1
   RUNG wire#powerrail
      Contact( #DATA.Elevateur.cmd.x_Stopper_down_manual )
   END_RUNG wire#w1
   RUNG wire#powerrail
      I_Contact( #x_en_auto )
      I_Contact( #x_en_demo )
   END_RUNG wire#w1
   // the same network as SCL:
   #_w1 := NOT #DATA.Elevateur.cmd.x_Stopper_down AND #Front_descendant_butee_elevateur;   // falling edge of #DATA.Elevateur.cmd.x_Stopper_down
   #Front_descendant_butee_elevateur := #DATA.Elevateur.cmd.x_Stopper_down;
   IF #DATA.Elevateur.cmd.x_Elevator_up THEN
       #DATA.Elevateur.status.x_Busy := TRUE;   // SR flip-flop
   END_IF;
   IF #_w1 OR #DATA.Elevateur.cmd.x_Stopper_down_manual OR (NOT #x_en_auto AND NOT #x_en_demo) THEN
       #DATA.Elevateur.status.x_Busy := FALSE;
   END_IF;
END_REGION

REGION Network 6: Gestion montee elevateur
   #IEC_Timer_0_Instance_1(IN := ((#x_en_auto AND (#DATA.Elevateur.status.x_Has_print_surface OR #x_All_stations_empty)) OR #x_en_demo) AND NOT #DATA.Elevateur.status.x_Fault AND NOT #x_defaut_externe AND #DATA.Elevateur.status.x_Pos_basse AND #DATA.Elevateur.status.x_Pres_palette AND NOT #DATA.Elevateur.cmd.x_Stopper_down AND NOT #DATA.Elevateur.status.x_Busy,   // TON
                           PT := T#250ms);
   IF #IEC_Timer_0_Instance_1.Q OR (#x_en_manu AND #DATA.Elevateur.cmd.x_Elevator_up_manual) THEN
       #DATA.Elevateur.cmd.x_Elevator_up := TRUE;   // SR flip-flop
   END_IF;
   IF #DATA.Elevateur.status.x_Pos_haute OR (#x_en_manu AND #DATA.Elevateur.cmd.x_Elevator_down_manual) OR #x_defaut_externe OR #DATA.Elevateur.status.x_Fault THEN
       #DATA.Elevateur.cmd.x_Elevator_up := FALSE;
   END_IF;
END_REGION

REGION Network 7: Gestion descente elevateur
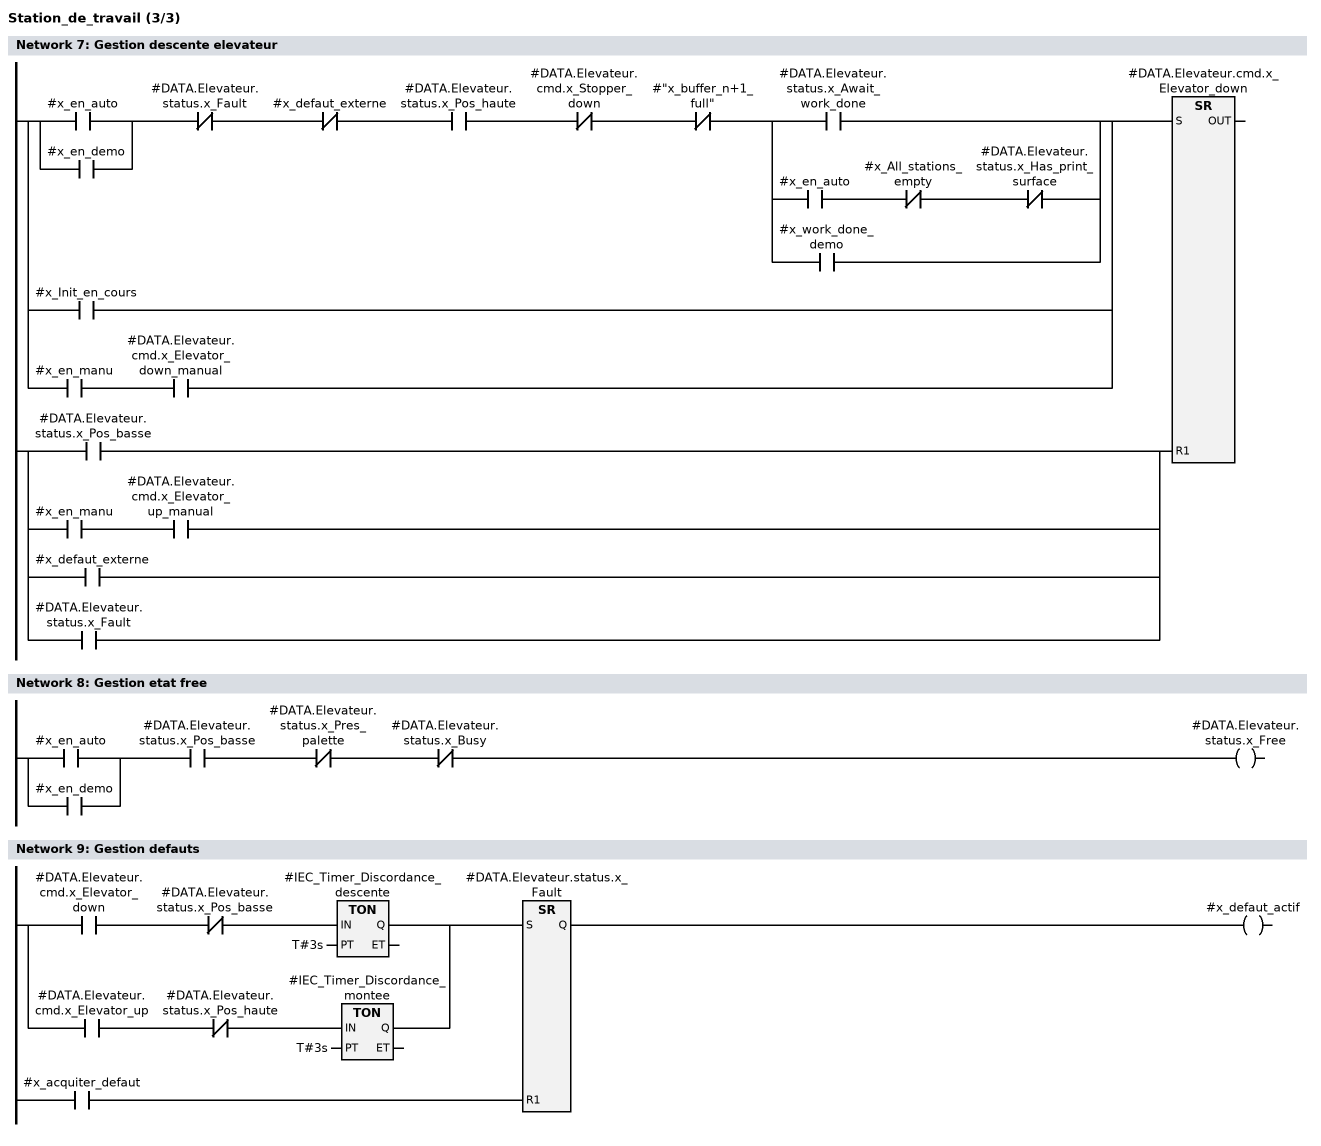
   RUNG wire#powerrail
      Contact( #x_en_auto )
      wire#w1
      I_Contact( #DATA.Elevateur.status.x_Fault )
      I_Contact( #x_defaut_externe )
      Contact( #DATA.Elevateur.status.x_Pos_haute )
      I_Contact( #DATA.Elevateur.cmd.x_Stopper_down )
      I_Contact( #"x_buffer_n+1_full" )
      wire#w2
      Contact( #DATA.Elevateur.status.x_Await_work_done )
      wire#w3
      S_SR(operand := #DATA.Elevateur.cmd.x_Elevator_down, r1 := wire#w4)
   END_RUNG
   RUNG wire#powerrail
      Contact( #x_en_demo )
   END_RUNG wire#w1
   RUNG wire#w2
      Contact( #x_en_auto )
      I_Contact( #x_All_stations_empty )
      I_Contact( #DATA.Elevateur.status.x_Has_print_surface )
   END_RUNG wire#w3
   RUNG wire#w2
      Contact( #x_work_done_demo )
   END_RUNG wire#w3
   RUNG wire#powerrail
      Contact( #x_Init_en_cours )
   END_RUNG wire#w3
   RUNG wire#powerrail
      Contact( #x_en_manu )
      Contact( #DATA.Elevateur.cmd.x_Elevator_down_manual )
   END_RUNG wire#w3
   RUNG wire#powerrail
      Contact( #DATA.Elevateur.status.x_Pos_basse )
   END_RUNG wire#w4
   RUNG wire#powerrail
      Contact( #x_en_manu )
      Contact( #DATA.Elevateur.cmd.x_Elevator_up_manual )
   END_RUNG wire#w4
   RUNG wire#powerrail
      Contact( #x_defaut_externe )
   END_RUNG wire#w4
   RUNG wire#powerrail
      Contact( #DATA.Elevateur.status.x_Fault )
   END_RUNG wire#w4
   // the same network as SCL:
   IF ((#x_en_auto OR #x_en_demo) AND NOT #DATA.Elevateur.status.x_Fault AND NOT #x_defaut_externe AND #DATA.Elevateur.status.x_Pos_haute AND NOT #DATA.Elevateur.cmd.x_Stopper_down AND NOT #"x_buffer_n+1_full" AND (#DATA.Elevateur.status.x_Await_work_done OR (#x_en_auto AND NOT #x_All_stations_empty AND NOT #DATA.Elevateur.status.x_Has_print_surface) OR #x_work_done_demo)) OR #x_Init_en_cours OR (#x_en_manu AND #DATA.Elevateur.cmd.x_Elevator_down_manual) THEN
       #DATA.Elevateur.cmd.x_Elevator_down := TRUE;   // SR flip-flop
   END_IF;
   IF #DATA.Elevateur.status.x_Pos_basse OR (#x_en_manu AND #DATA.Elevateur.cmd.x_Elevator_up_manual) OR #x_defaut_externe OR #DATA.Elevateur.status.x_Fault THEN
       #DATA.Elevateur.cmd.x_Elevator_down := FALSE;
   END_IF;
END_REGION

REGION Network 8: Gestion etat free
   RUNG wire#powerrail
      Contact( #x_en_auto )
      wire#w1
      Contact( #DATA.Elevateur.status.x_Pos_basse )
      I_Contact( #DATA.Elevateur.status.x_Pres_palette )
      I_Contact( #DATA.Elevateur.status.x_Busy )
      Coil( #DATA.Elevateur.status.x_Free )
   END_RUNG
   RUNG wire#powerrail
      Contact( #x_en_demo )
   END_RUNG wire#w1
   // the same network as SCL:
   #DATA.Elevateur.status.x_Free := (#x_en_auto OR #x_en_demo) AND #DATA.Elevateur.status.x_Pos_basse AND NOT #DATA.Elevateur.status.x_Pres_palette AND NOT #DATA.Elevateur.status.x_Busy;
END_REGION

REGION Network 9: Gestion defauts
   #IEC_Timer_Discordance_descente(IN := #DATA.Elevateur.cmd.x_Elevator_down AND NOT #DATA.Elevateur.status.x_Pos_basse,   // TON
                           PT := T#3s);
   #IEC_Timer_Discordance_montee(IN := #DATA.Elevateur.cmd.x_Elevator_up AND NOT #DATA.Elevateur.status.x_Pos_haute,   // TON
                           PT := T#3s);
   IF #IEC_Timer_Discordance_descente.Q OR #IEC_Timer_Discordance_montee.Q THEN
       #DATA.Elevateur.status.x_Fault := TRUE;   // SR flip-flop
   END_IF;
   IF #x_acquiter_defaut THEN #DATA.Elevateur.status.x_Fault := FALSE; END_IF;
   #x_defaut_actif := #DATA.Elevateur.status.x_Fault;
END_REGION
END_FUNCTION_BLOCK

// folder: 200_Generateur_Alarmes

FUNCTION_BLOCK "Create_Alarm"   // FB1, LAD
{ S7_Optimized_Access := 'TRUE' }
VERSION : 0.1
   VAR_INPUT
      x_Alarm_input : Bool;
      str_Tag : String;
      str_Alarm_text : String;
   END_VAR
   VAR_OUTPUT
      x_Error : Bool;
   END_VAR
   VAR
      Program_Alarm_1 : Program_Alarm;
   END_VAR
   VAR_TEMP
      w_Status : Word;
   END_VAR
BEGIN

REGION Network 1
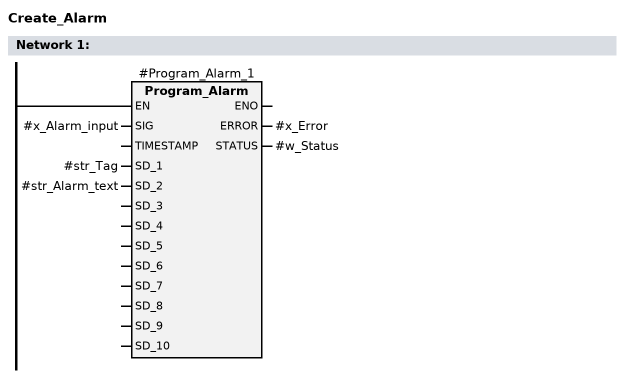
   #Program_Alarm_1(SIG := #x_Alarm_input,   // Program_Alarm
                    SD_1 := #str_Tag,
                    SD_2 := #str_Alarm_text,
                    Error => #x_Error,
                    Status => #w_Status);
END_REGION
END_FUNCTION_BLOCK

// folder: 3_Controle vision

FUNCTION_BLOCK "FIFO"   // FB12, LAD
{ S7_Optimized_Access := 'TRUE' }
VERSION : 0.1
   VAR_INPUT
      I : Int;
   END_VAR
   VAR_OUTPUT
      O : Int;
   END_VAR
   VAR
      Float_1 : Int;
      Float_2 : Int;
      Float_3 : Int;
   END_VAR
BEGIN

REGION Network 1
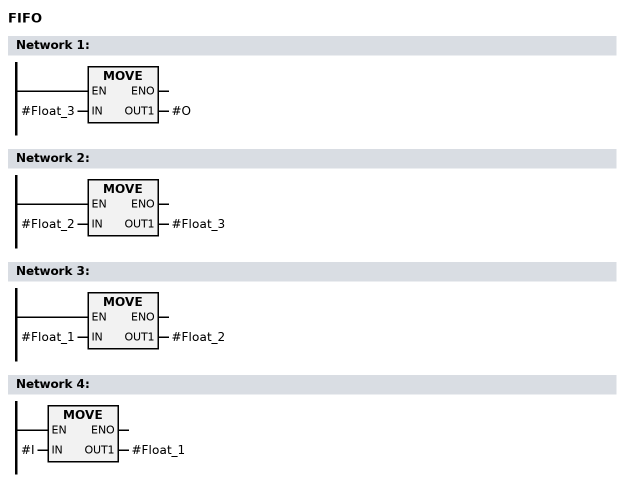
   RUNG wire#powerrail
      Move(in := #Float_3, out1 => #O)
   END_RUNG
   // the same network as SCL:
   #O := #Float_3;
END_REGION

REGION Network 2
   RUNG wire#powerrail
      Move(in := #Float_2, out1 => #Float_3)
   END_RUNG
   // the same network as SCL:
   #Float_3 := #Float_2;
END_REGION

REGION Network 3
   RUNG wire#powerrail
      Move(in := #Float_1, out1 => #Float_2)
   END_RUNG
   // the same network as SCL:
   #Float_2 := #Float_1;
END_REGION

REGION Network 4
   RUNG wire#powerrail
      Move(in := #I, out1 => #Float_1)
   END_RUNG
   // the same network as SCL:
   #Float_1 := #I;
END_REGION
END_FUNCTION_BLOCK

FUNCTION_BLOCK "31_Keyence_Camera"   // FB13, LAD
{ S7_Optimized_Access := 'TRUE' }
VERSION : 0.1
BEGIN
END_FUNCTION_BLOCK

FUNCTION_BLOCK "32_Cmd_porte_vision"   // FB14, LAD
{ S7_Optimized_Access := 'TRUE' }
VERSION : 0.1
   VAR
      x_ouverture_porte_vision : Bool;
      x_fermeture_porte_vision : Bool;
      x_Ouverture_porte_manu : Bool;
      x_Fermeture_porte_manu : Bool;
   END_VAR
BEGIN

REGION Network 1: Ouverture porte vision
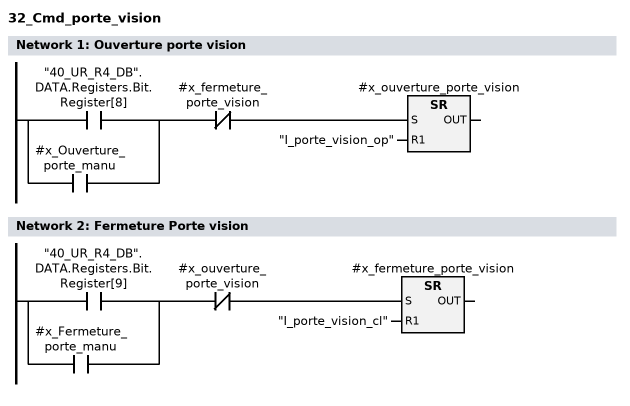
   RUNG wire#powerrail
      Contact( "40_UR_R4_DB".DATA.Registers.Bit.Register[8] )
      wire#w1
      I_Contact( #x_fermeture_porte_vision )
      S_SR(operand := #x_ouverture_porte_vision, r1 := "I_porte_vision_op")
   END_RUNG
   RUNG wire#powerrail
      Contact( #x_Ouverture_porte_manu )
   END_RUNG wire#w1
   // the same network as SCL:
   IF ("40_UR_R4_DB".DATA.Registers.Bit.Register[8] OR #x_Ouverture_porte_manu) AND NOT #x_fermeture_porte_vision THEN
       #x_ouverture_porte_vision := TRUE;   // SR flip-flop
   END_IF;
   IF "I_porte_vision_op" THEN #x_ouverture_porte_vision := FALSE; END_IF;
END_REGION

REGION Network 2: Fermeture Porte vision
   RUNG wire#powerrail
      Contact( "40_UR_R4_DB".DATA.Registers.Bit.Register[9] )
      wire#w1
      I_Contact( #x_ouverture_porte_vision )
      S_SR(operand := #x_fermeture_porte_vision, r1 := "I_porte_vision_cl")
   END_RUNG
   RUNG wire#powerrail
      Contact( #x_Fermeture_porte_manu )
   END_RUNG wire#w1
   // the same network as SCL:
   IF ("40_UR_R4_DB".DATA.Registers.Bit.Register[9] OR #x_Fermeture_porte_manu) AND NOT #x_ouverture_porte_vision THEN
       #x_fermeture_porte_vision := TRUE;   // SR flip-flop
   END_IF;
   IF "I_porte_vision_cl" THEN #x_fermeture_porte_vision := FALSE; END_IF;
END_REGION
END_FUNCTION_BLOCK

FUNCTION "Controle_vision_provisoire" : Void   // FC16, LAD
{ S7_Optimized_Access := 'TRUE' }
VERSION : 0.1
   VAR_TEMP   // added for the SCL form of the ladder/FBD networks
      _w1 : Bool;
   END_VAR
BEGIN

REGION Network 1: Envoi trigger
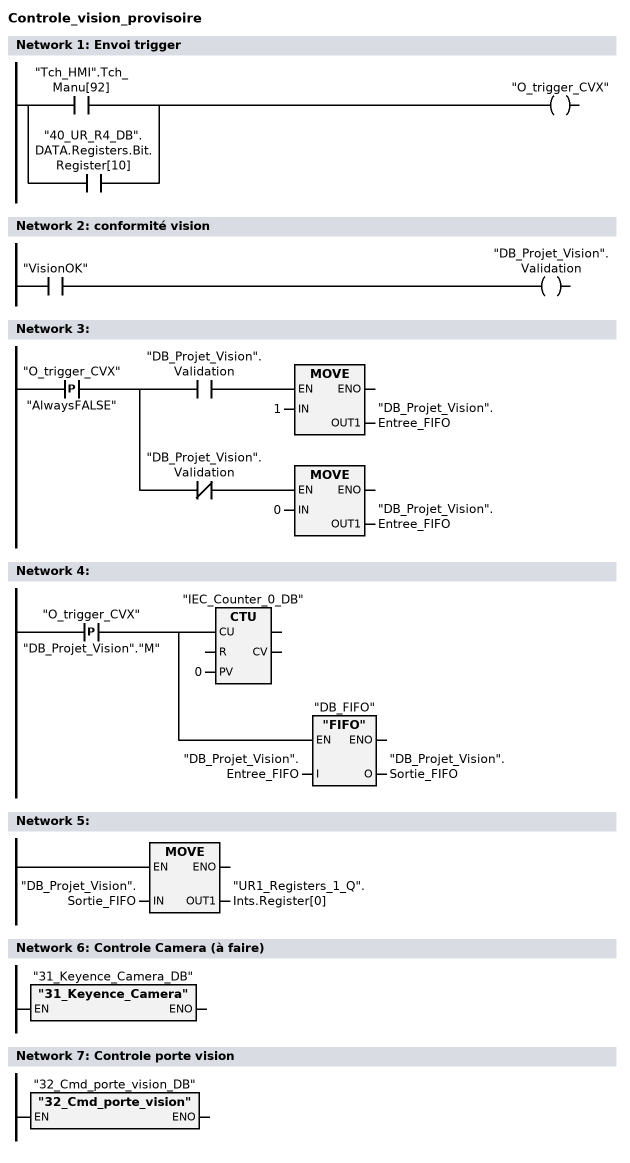
   RUNG wire#powerrail
      Contact( "Tch_HMI".Tch_Manu[92] )
      wire#w1
      Coil( "O_trigger_CVX" )
   END_RUNG
   RUNG wire#powerrail
      Contact( "40_UR_R4_DB".DATA.Registers.Bit.Register[10] )
   END_RUNG wire#w1
   // the same network as SCL:
   "O_trigger_CVX" := "Tch_HMI".Tch_Manu[92] OR "40_UR_R4_DB".DATA.Registers.Bit.Register[10];
END_REGION

REGION Network 2: conformité vision
   RUNG wire#powerrail
      Contact( "VisionOK" )
      Coil( "DB_Projet_Vision".Validation )
   END_RUNG
   // the same network as SCL:
   "DB_Projet_Vision".Validation := "VisionOK";
END_REGION

REGION Network 3
   RUNG wire#powerrail
      P_Contact(operand := "O_trigger_CVX", bit := "AlwaysFALSE")
      wire#w1
      Contact( "DB_Projet_Vision".Validation )
      Move(in := 1, out1 => "DB_Projet_Vision".Entree_FIFO)
   END_RUNG
   RUNG wire#w1
      I_Contact( "DB_Projet_Vision".Validation )
      Move(in := 0, out1 => "DB_Projet_Vision".Entree_FIFO)
   END_RUNG
   // the same network as SCL:
   #_w1 := "O_trigger_CVX" AND NOT "AlwaysFALSE";   // rising edge of "O_trigger_CVX"
   "AlwaysFALSE" := "O_trigger_CVX";
   IF #_w1 AND "DB_Projet_Vision".Validation THEN "DB_Projet_Vision".Entree_FIFO := 1; END_IF;
   IF #_w1 AND NOT "DB_Projet_Vision".Validation THEN "DB_Projet_Vision".Entree_FIFO := 0; END_IF;
END_REGION

REGION Network 4
   #_w1 := "O_trigger_CVX" AND NOT "DB_Projet_Vision"."M";   // rising edge of "O_trigger_CVX"
   "DB_Projet_Vision"."M" := "O_trigger_CVX";
   "IEC_Counter_0_DB".CTU(CU := #_w1, PV := 0);
   IF #_w1 THEN
       "DB_FIFO"(I := "DB_Projet_Vision".Entree_FIFO, O => "DB_Projet_Vision".Sortie_FIFO);   // "FIFO"
   END_IF;
END_REGION

REGION Network 5
   RUNG wire#powerrail
      Move(in := "DB_Projet_Vision".Sortie_FIFO, out1 => "UR1_Registers_1_Q".Ints.Register[0])
   END_RUNG
   // the same network as SCL:
   "UR1_Registers_1_Q".Ints.Register[0] := "DB_Projet_Vision".Sortie_FIFO;
END_REGION

REGION Network 6: Controle Camera (à faire)
   RUNG wire#powerrail
      "31_Keyence_Camera_DB"()
   END_RUNG
   // the same network as SCL:
   "31_Keyence_Camera_DB"();   // "31_Keyence_Camera"
END_REGION

REGION Network 7: Controle porte vision
   RUNG wire#powerrail
      "32_Cmd_porte_vision_DB"()
   END_RUNG
   // the same network as SCL:
   "32_Cmd_porte_vision_DB"();   // "32_Cmd_porte_vision"
END_REGION
END_FUNCTION

// folder: 4_UR10_R4

FUNCTION_BLOCK "40_UR_R4"   // FB4, LAD
{ S7_Optimized_Access := 'TRUE' }
VERSION : 0.1
   VAR
      DATA : "UR_Cobot";
      DmdEcritureModbusAGV2 : Bool;
   END_VAR
   // // DATA.Registers_Out_1.Bits.Register[0] : Work done imprimante 1
   // // DATA.Registers_Out_1.Bits.Register[1] : Work done imprimante 2
   // // DATA.Registers_Out_1.Bits.Register[2] : Work done imprimante 3
   // // DATA.Registers_Out_1.Bits.Register[3] : Work done imprimante 4
   // // DATA.Registers_Out_1.Bits.Register[4] : Work done imprimante 5
   // // DATA.Registers_Out_1.Bits.Register[5] : Work done imprimante 6
   // // DATA.Registers_Out_1.Bits.Register[6] : Work done imprimante 7
   // // DATA.Registers_Out_1.Bits.Register[7] : Work done imprimante 8
   // // DATA.Registers_Out_1.Bits.Register[8] : Poste 1 Dispo
   // // DATA.Registers_Out_1.Bits.Register[9] : Poste 2 Dispo
   // // DATA.Registers_Out_1.Bits.Register[10] : Poste 3 Dispo
   // // DATA.Registers_Out_1.Bits.Register[11] : Poste 4 Dispo
   // // DATA.Registers_Out_1.Bits.Register[12] : Poste 5 Dispo
   // // DATA.Registers_Out_1.Bits.Register[13] : Poste 6 Dispo
   // // DATA.Registers_Out_1.Bits.Register[14] : Poste 7 Dispo
   // // DATA.Registers_Out_2.Bits.Register[0] : Demande Init
   // // DATA.Registers_Out_2.Bits.Register[1] : EnCycleAuto
   // // DATA.Registers_Out_2.Bits.Register[2] : EnCycleDemo
   // // DATA.Registers_Out_2.Bits.Register[3] : PauseProgPLC
   // // DATA.Registers_Out_2.Bits.Register[4] : StopProgPLC
   // // DATA.Registers_Out_2.Bits.Register[5] : StartProgPLC (demarrage boucle Main)
   // // DATA.Registers_Out_2.Bits.Register[6] : Initialisation auto après AU
   // // DATA.Registers.Bit.Register[1] : WorkDoneP1
   // // DATA.Registers.Bit.Register[2] : WorkDoneP2
   // // DATA.Registers.Bit.Register[3] : WorkDoneP3
   // // DATA.Registers.Bit.Register[4] : WorkDoneP4
   // // DATA.Registers.Bit.Register[5] : WorkDoneP5
   // // DATA.Registers.Bit.Register[6] : WorkDoneP6
   // // DATA.Registers.Bit.Register[7] : WorkDoneP7
   // // DATA.Registers.Bit.Register[8] : Dmd Ouverture porte Vision
   // // DATA.Registers.Bit.Register[9] : Dmd Fermeture porte Vision
   // // DATA.Registers.Bit.Register[10] : Trigger Vision
   // // DATA.Registers_Out_2.Bits.Register[7] : InitRequired
   // // DATA.Registers.Bit.Register[0] : IsInitialized
   // // DATA.Registers_Out_2.Bits.Register[8] : UnpauseProgPLC
   // // DATA.Registers_Out_1.Bits.Register[15] : Porte Vision Open
   // // DATA.Registers_Out_1.Bits.Register[16] : Porte Vision fermee
   // // DATA.Registers_Out_1.Bits.Register[17] : Vision prete
   // // DATA.Registers_Out_1.Bits.Register[18] : ColisVideDispo
   // // DATA.Registers_Out_1.Bits.Register[19] : CouvercleRecuperee
   // // DATA.Registers.Bit.Register[11] : FinDeposeColis
   // // DATA.Registers.Bit.Register[12] : PosRecupCouvercle
   // // DATA.Registers_Out_2.Bits.Register[9] : VisionOK2
   // // DATA.Registers_Out_1.Bits.Register[20] : VisionOk
BEGIN

REGION Network 1: Init Required?
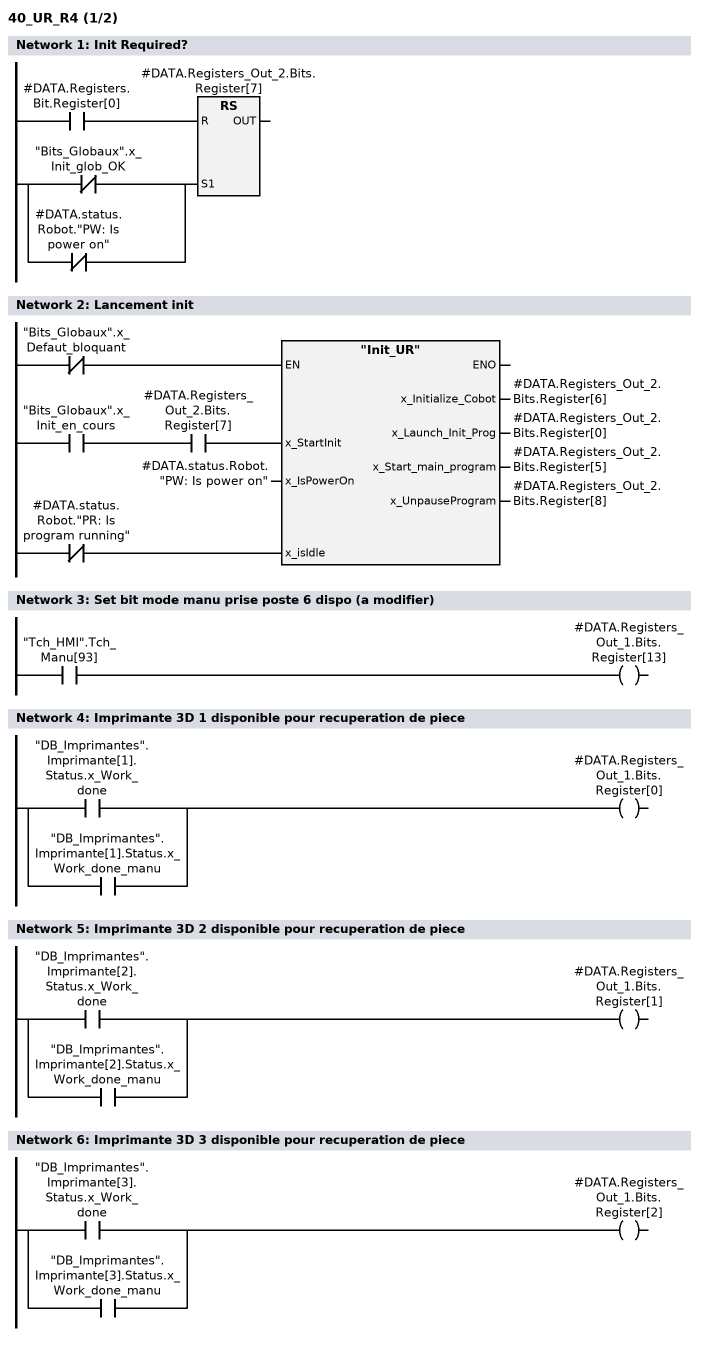
   RUNG wire#powerrail
      Contact( #DATA.Registers.Bit.Register[0] )
      S_RS(operand := #DATA.Registers_Out_2.Bits.Register[7], s1 := wire#w1)
   END_RUNG
   RUNG wire#powerrail
      I_Contact( "Bits_Globaux".x_Init_glob_OK )
   END_RUNG wire#w1
   RUNG wire#powerrail
      I_Contact( #DATA.status.Robot."PW: Is power on" )
   END_RUNG wire#w1
   // the same network as SCL:
   IF #DATA.Registers.Bit.Register[0] THEN
       #DATA.Registers_Out_2.Bits.Register[7] := FALSE;   // RS flip-flop
   END_IF;
   IF NOT "Bits_Globaux".x_Init_glob_OK OR NOT #DATA.status.Robot."PW: Is power on" THEN
       #DATA.Registers_Out_2.Bits.Register[7] := TRUE;
   END_IF;
END_REGION

REGION Network 2: Lancement init
   RUNG wire#powerrail
      I_Contact( "Bits_Globaux".x_Defaut_bloquant )
      "Init_UR"(x_StartInit := wire#w1, x_isIdle := wire#w2, x_IsPowerOn := #DATA.status.Robot."PW: Is power on", x_Initialize_Cobot => #DATA.Registers_Out_2.Bits.Register[6], x_Launch_Init_Prog => #DATA.Registers_Out_2.Bits.Register[0], x_Start_main_program => #DATA.Registers_Out_2.Bits.Register[5], x_UnpauseProgram => #DATA.Registers_Out_2.Bits.Register[8])
   END_RUNG
   RUNG wire#powerrail
      Contact( "Bits_Globaux".x_Init_en_cours )
      Contact( #DATA.Registers_Out_2.Bits.Register[7] )
   END_RUNG wire#w1
   RUNG wire#powerrail
      I_Contact( #DATA.status.Robot."PR: Is program running" )
   END_RUNG wire#w2
   // the same network as SCL:
   IF NOT "Bits_Globaux".x_Defaut_bloquant THEN
       "Init_UR"(x_StartInit := "Bits_Globaux".x_Init_en_cours AND #DATA.Registers_Out_2.Bits.Register[7],
                 x_IsPowerOn := #DATA.status.Robot."PW: Is power on",
                 x_isIdle := NOT #DATA.status.Robot."PR: Is program running",
                 x_Initialize_Cobot => #DATA.Registers_Out_2.Bits.Register[6],
                 x_Launch_Init_Prog => #DATA.Registers_Out_2.Bits.Register[0],
                 x_Start_main_program => #DATA.Registers_Out_2.Bits.Register[5],
                 x_UnpauseProgram => #DATA.Registers_Out_2.Bits.Register[8]);
   END_IF;
END_REGION

REGION Network 3: Set bit mode manu prise poste 6 dispo (a modifier)
   RUNG wire#powerrail
      Contact( "Tch_HMI".Tch_Manu[93] )
      Coil( #DATA.Registers_Out_1.Bits.Register[13] )
   END_RUNG
   // the same network as SCL:
   #DATA.Registers_Out_1.Bits.Register[13] := "Tch_HMI".Tch_Manu[93];
END_REGION

REGION Network 4: Imprimante 3D 1 disponible pour recuperation de piece
   RUNG wire#powerrail
      Contact( "DB_Imprimantes".Imprimante[1].Status.x_Work_done )
      wire#w1
      Coil( #DATA.Registers_Out_1.Bits.Register[0] )
   END_RUNG
   RUNG wire#powerrail
      Contact( "DB_Imprimantes".Imprimante[1].Status.x_Work_done_manu )
   END_RUNG wire#w1
   // the same network as SCL:
   #DATA.Registers_Out_1.Bits.Register[0] := "DB_Imprimantes".Imprimante[1].Status.x_Work_done OR "DB_Imprimantes".Imprimante[1].Status.x_Work_done_manu;
END_REGION

REGION Network 5: Imprimante 3D 2 disponible pour recuperation de piece
   RUNG wire#powerrail
      Contact( "DB_Imprimantes".Imprimante[2].Status.x_Work_done )
      wire#w1
      Coil( #DATA.Registers_Out_1.Bits.Register[1] )
   END_RUNG
   RUNG wire#powerrail
      Contact( "DB_Imprimantes".Imprimante[2].Status.x_Work_done_manu )
   END_RUNG wire#w1
   // the same network as SCL:
   #DATA.Registers_Out_1.Bits.Register[1] := "DB_Imprimantes".Imprimante[2].Status.x_Work_done OR "DB_Imprimantes".Imprimante[2].Status.x_Work_done_manu;
END_REGION

REGION Network 6: Imprimante 3D 3 disponible pour recuperation de piece
   RUNG wire#powerrail
      Contact( "DB_Imprimantes".Imprimante[3].Status.x_Work_done )
      wire#w1
      Coil( #DATA.Registers_Out_1.Bits.Register[2] )
   END_RUNG
   RUNG wire#powerrail
      Contact( "DB_Imprimantes".Imprimante[3].Status.x_Work_done_manu )
   END_RUNG wire#w1
   // the same network as SCL:
   #DATA.Registers_Out_1.Bits.Register[2] := "DB_Imprimantes".Imprimante[3].Status.x_Work_done OR "DB_Imprimantes".Imprimante[3].Status.x_Work_done_manu;
END_REGION

REGION Network 7: Imprimante 3D 4 disponible pour recuperation de piece
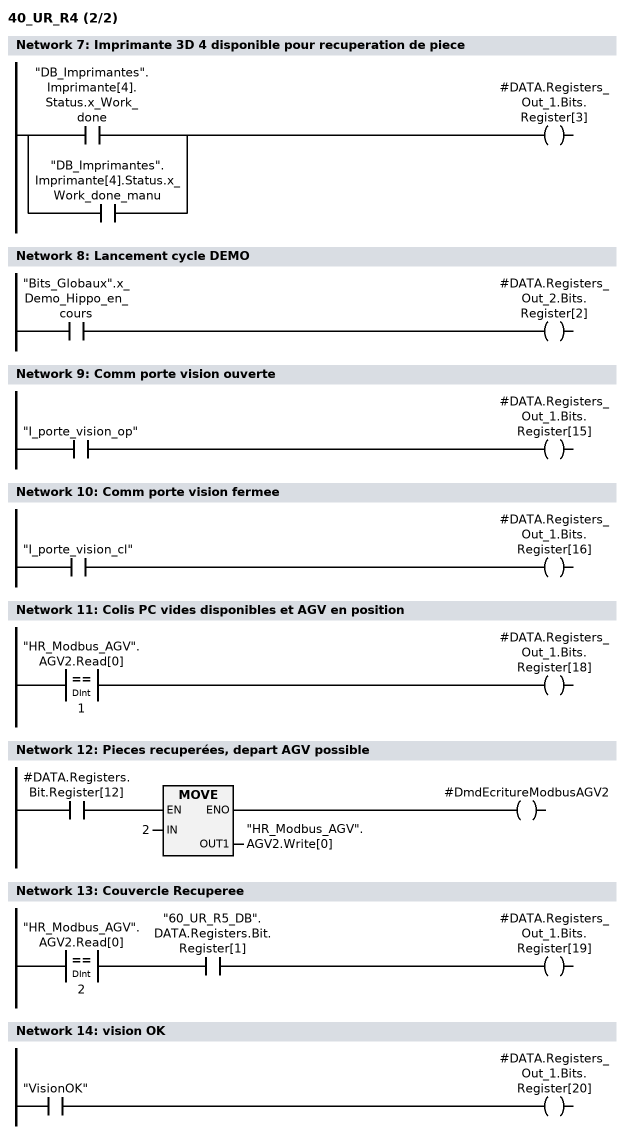
   RUNG wire#powerrail
      Contact( "DB_Imprimantes".Imprimante[4].Status.x_Work_done )
      wire#w1
      Coil( #DATA.Registers_Out_1.Bits.Register[3] )
   END_RUNG
   RUNG wire#powerrail
      Contact( "DB_Imprimantes".Imprimante[4].Status.x_Work_done_manu )
   END_RUNG wire#w1
   // the same network as SCL:
   #DATA.Registers_Out_1.Bits.Register[3] := "DB_Imprimantes".Imprimante[4].Status.x_Work_done OR "DB_Imprimantes".Imprimante[4].Status.x_Work_done_manu;
END_REGION

REGION Network 8: Lancement cycle DEMO
   RUNG wire#powerrail
      Contact( "Bits_Globaux".x_Demo_Hippo_en_cours )
      Coil( #DATA.Registers_Out_2.Bits.Register[2] )
   END_RUNG
   // the same network as SCL:
   #DATA.Registers_Out_2.Bits.Register[2] := "Bits_Globaux".x_Demo_Hippo_en_cours;
END_REGION

REGION Network 9: Comm porte vision ouverte
   RUNG wire#powerrail
      Contact( "I_porte_vision_op" )
      Coil( #DATA.Registers_Out_1.Bits.Register[15] )
   END_RUNG
   // the same network as SCL:
   #DATA.Registers_Out_1.Bits.Register[15] := "I_porte_vision_op";
END_REGION

REGION Network 10: Comm porte vision fermee
   RUNG wire#powerrail
      Contact( "I_porte_vision_cl" )
      Coil( #DATA.Registers_Out_1.Bits.Register[16] )
   END_RUNG
   // the same network as SCL:
   #DATA.Registers_Out_1.Bits.Register[16] := "I_porte_vision_cl";
END_REGION

REGION Network 11: Colis PC vides disponibles et AGV en position
   RUNG wire#powerrail
      { S7_Templates := "SrcType := DInt" } EQ_Contact(in1 := "HR_Modbus_AGV".AGV2.Read[0], in2 := 1)
      Coil( #DATA.Registers_Out_1.Bits.Register[18] )
   END_RUNG
   // the same network as SCL:
   #DATA.Registers_Out_1.Bits.Register[18] := "HR_Modbus_AGV".AGV2.Read[0] = 1;
END_REGION

REGION Network 12: Pieces recuperées, depart AGV possible
   RUNG wire#powerrail
      Contact( #DATA.Registers.Bit.Register[12] )
      Move(in := 2, out1 => "HR_Modbus_AGV".AGV2.Write[0])
      Coil( #DmdEcritureModbusAGV2 )
   END_RUNG
   // the same network as SCL:
   IF #DATA.Registers.Bit.Register[12] THEN "HR_Modbus_AGV".AGV2.Write[0] := 2; END_IF;
   #DmdEcritureModbusAGV2 := #DATA.Registers.Bit.Register[12];
END_REGION

REGION Network 13: Couvercle Recuperee
   RUNG wire#powerrail
      { S7_Templates := "SrcType := DInt" } EQ_Contact(in1 := "HR_Modbus_AGV".AGV2.Read[0], in2 := 2)
      Contact( "60_UR_R5_DB".DATA.Registers.Bit.Register[1] )
      Coil( #DATA.Registers_Out_1.Bits.Register[19] )
   END_RUNG
   // the same network as SCL:
   #DATA.Registers_Out_1.Bits.Register[19] := ("HR_Modbus_AGV".AGV2.Read[0] = 2) AND "60_UR_R5_DB".DATA.Registers.Bit.Register[1];
END_REGION

REGION Network 14: vision OK
   RUNG wire#powerrail
      Contact( "VisionOK" )
      Coil( #DATA.Registers_Out_1.Bits.Register[20] )
   END_RUNG
   // the same network as SCL:
   #DATA.Registers_Out_1.Bits.Register[20] := "VisionOK";
END_REGION
END_FUNCTION_BLOCK

FUNCTION "Init_UR" : Void   // FC20, LAD
{ S7_Optimized_Access := 'TRUE' }
VERSION : 0.1
   VAR_INPUT
      x_StartInit : Bool;
      x_IsPowerOn : Bool;
      x_isIdle : Bool;
   END_VAR
   VAR_OUTPUT
      x_Initialize_Cobot : Bool;
      x_Launch_Init_Prog : Bool;
      x_Start_main_program : Bool;
      x_UnpauseProgram : Bool;
   END_VAR
BEGIN

REGION Network 1: Verification etat robot et lancement initialisation avec deblocage des freins
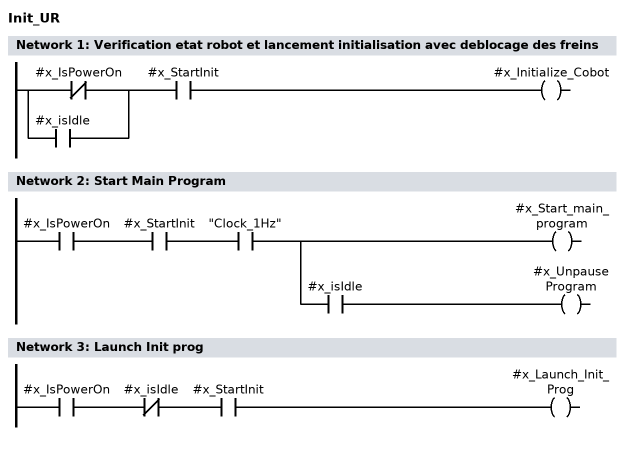
   RUNG wire#powerrail
      I_Contact( #x_IsPowerOn )
      wire#w1
      Contact( #x_StartInit )
      Coil( #x_Initialize_Cobot )
   END_RUNG
   RUNG wire#powerrail
      Contact( #x_isIdle )
   END_RUNG wire#w1
   // the same network as SCL:
   #x_Initialize_Cobot := (NOT #x_IsPowerOn OR #x_isIdle) AND #x_StartInit;
END_REGION

REGION Network 2: Start Main Program
   RUNG wire#powerrail
      Contact( #x_IsPowerOn )
      Contact( #x_StartInit )
      Contact( "Clock_1Hz" )
      wire#w1
      Coil( #x_Start_main_program )
   END_RUNG
   RUNG wire#w1
      Contact( #x_isIdle )
      Coil( #x_UnpauseProgram )
   END_RUNG
   // the same network as SCL:
   #x_Start_main_program := #x_IsPowerOn AND #x_StartInit AND "Clock_1Hz";
   #x_UnpauseProgram := #x_Start_main_program AND #x_isIdle;
END_REGION

REGION Network 3: Launch Init prog
   RUNG wire#powerrail
      Contact( #x_IsPowerOn )
      I_Contact( #x_isIdle )
      Contact( #x_StartInit )
      Coil( #x_Launch_Init_Prog )
   END_RUNG
   // the same network as SCL:
   #x_Launch_Init_Prog := #x_IsPowerOn AND NOT #x_isIdle AND #x_StartInit;
END_REGION
END_FUNCTION

// folder: 5-Cellule_conditionnement

FUNCTION "50_Cellule_de_conditionnement" : Void   // FC13, LAD
{ S7_Optimized_Access := 'TRUE' }
VERSION : 0.1
BEGIN

REGION Network 1: Programme FANUC R1 (ajouter UDT de type Robot FANUC)
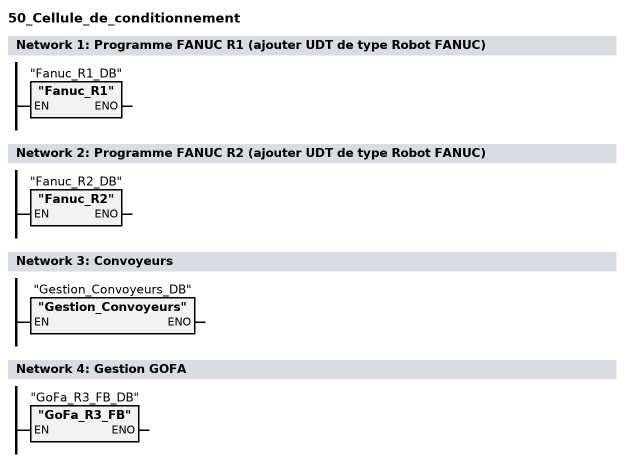
   RUNG wire#powerrail
      "Fanuc_R1_DB"()
   END_RUNG
   // the same network as SCL:
   "Fanuc_R1_DB"();   // "Fanuc_R1"
END_REGION

REGION Network 2: Programme FANUC R2 (ajouter UDT de type Robot FANUC)
   RUNG wire#powerrail
      "Fanuc_R2_DB"()
   END_RUNG
   // the same network as SCL:
   "Fanuc_R2_DB"();   // "Fanuc_R2"
END_REGION

REGION Network 3: Convoyeurs
   RUNG wire#powerrail
      "Gestion_Convoyeurs_DB"()
   END_RUNG
   // the same network as SCL:
   "Gestion_Convoyeurs_DB"();   // "Gestion_Convoyeurs"
END_REGION

REGION Network 4: Gestion GOFA
   RUNG wire#powerrail
      "GoFa_R3_FB_DB"()
   END_RUNG
   // the same network as SCL:
   "GoFa_R3_FB_DB"();   // "GoFa_R3_FB"
END_REGION
END_FUNCTION

// folder: 5-Cellule_conditionnement/Convoyeurs

FUNCTION_BLOCK "Convoyeur_conditionnement"   // FB2, LAD
TITLE = Controle convoyeur avec variateur zone de conditionnement
{ S7_Optimized_Access := 'TRUE' }
VERSION : 0.1
   VAR_INPUT
      Cpt_entree : Bool;
      Cpt_milieu : Bool;
      Cpt_fin : Bool;
      DefautExterneActif : Bool;
      AvecSAS : Bool;   // 0 ou 1
      "Vitesse MANU" : Int;
      "Vitesse AUTO" : Int;
      Ack_defaut : Bool;
      Rearmement : Bool;
      MarcheMoteurAuto : Bool;
      MarcheMoteurManu : Bool;
      DelaiArretMoteur : Time;   // en ms
      PorteOuverte : Bool;   // Arret moteur si porte ouverte
      Dmd_Arret : Bool;
      InversionSens : Bool;
   END_VAR
   VAR_OUTPUT
      DefautVariateur : Bool;
   END_VAR
   VAR_IN_OUT
      DB_Variateur : "Var_G120C_data";
   END_VAR
   VAR
      DB_Retard_arret_moteur : TON_TIME;
      Ft_montant_cpt : Bool;
   END_VAR
   VAR_TEMP
      ResultNorm_sp : Real;
      ResultScale_sp : Int;
   END_VAR
   VAR_TEMP   // added for the SCL form of the ladder/FBD networks
      _w1 : Bool;
   END_VAR
BEGIN

REGION Network 1: Activation pilotage par API
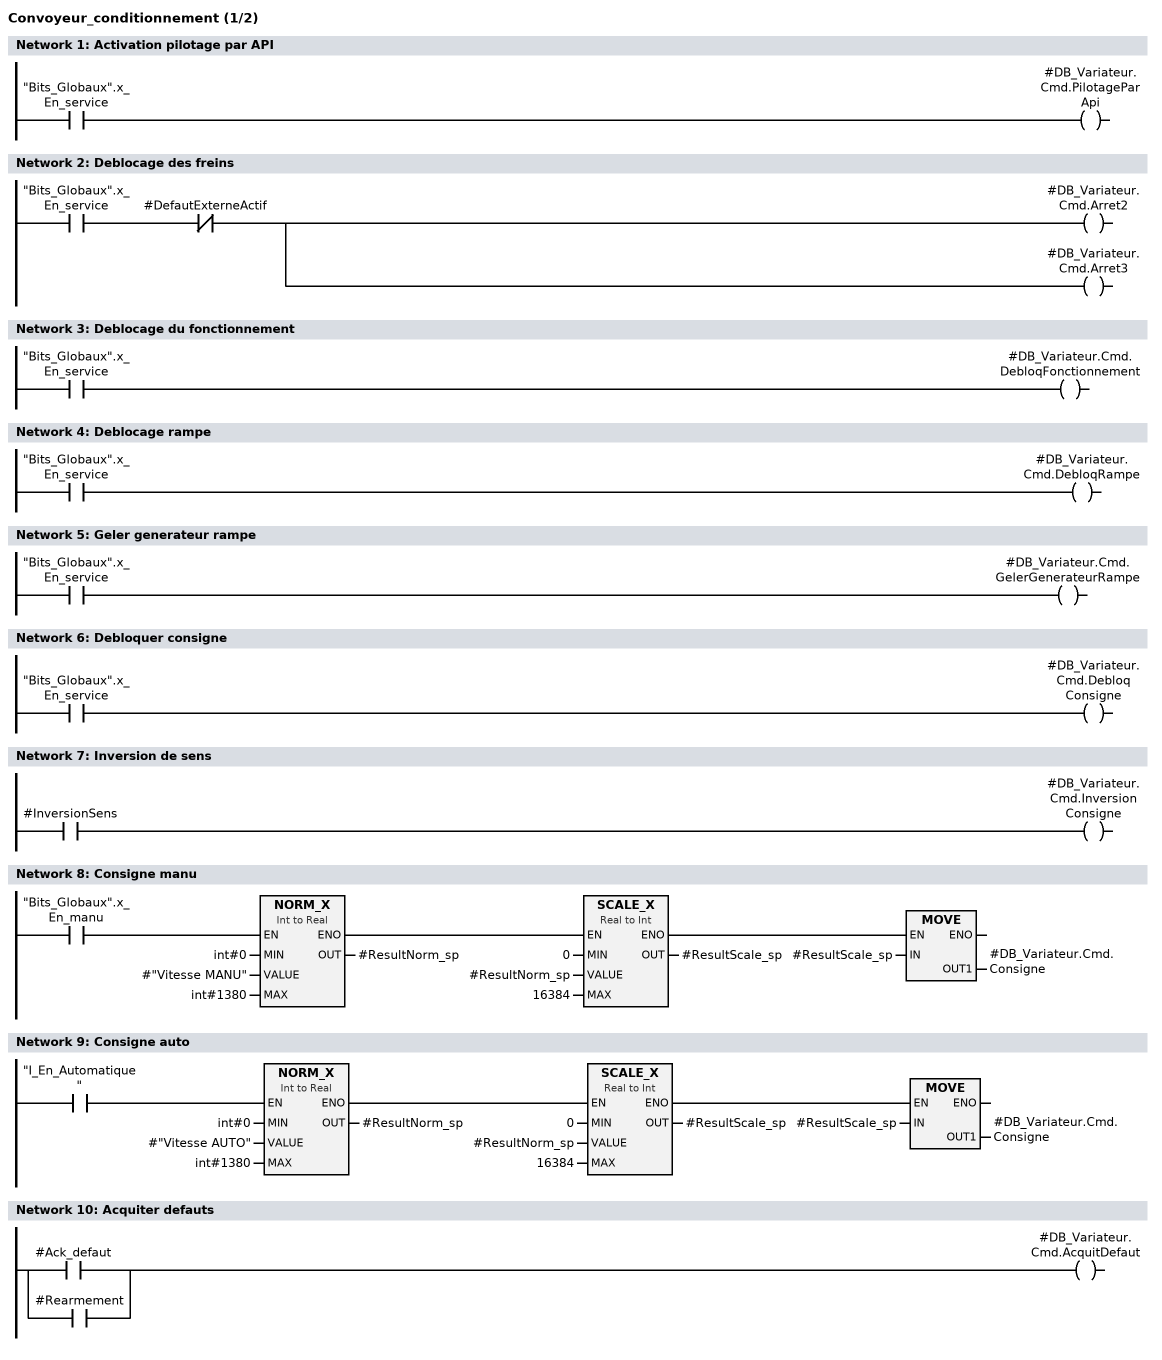
   RUNG wire#powerrail
      Contact( "Bits_Globaux".x_En_service )
      Coil( #DB_Variateur.Cmd.PilotageParApi )
   END_RUNG
   // the same network as SCL:
   #DB_Variateur.Cmd.PilotageParApi := "Bits_Globaux".x_En_service;
END_REGION

REGION Network 2: Deblocage des freins
   RUNG wire#powerrail
      Contact( "Bits_Globaux".x_En_service )
      I_Contact( #DefautExterneActif )
      wire#w1
      Coil( #DB_Variateur.Cmd.Arret2 )
   END_RUNG
   RUNG wire#w1
      Coil( #DB_Variateur.Cmd.Arret3 )
   END_RUNG
   // the same network as SCL:
   #DB_Variateur.Cmd.Arret2 := "Bits_Globaux".x_En_service AND NOT #DefautExterneActif;
   #DB_Variateur.Cmd.Arret3 := #DB_Variateur.Cmd.Arret2;
END_REGION

REGION Network 3: Deblocage du fonctionnement
   RUNG wire#powerrail
      Contact( "Bits_Globaux".x_En_service )
      Coil( #DB_Variateur.Cmd.DebloqFonctionnement )
   END_RUNG
   // the same network as SCL:
   #DB_Variateur.Cmd.DebloqFonctionnement := "Bits_Globaux".x_En_service;
END_REGION

REGION Network 4: Deblocage rampe
   RUNG wire#powerrail
      Contact( "Bits_Globaux".x_En_service )
      Coil( #DB_Variateur.Cmd.DebloqRampe )
   END_RUNG
   // the same network as SCL:
   #DB_Variateur.Cmd.DebloqRampe := "Bits_Globaux".x_En_service;
END_REGION

REGION Network 5: Geler generateur rampe
   RUNG wire#powerrail
      Contact( "Bits_Globaux".x_En_service )
      Coil( #DB_Variateur.Cmd.GelerGenerateurRampe )
   END_RUNG
   // the same network as SCL:
   #DB_Variateur.Cmd.GelerGenerateurRampe := "Bits_Globaux".x_En_service;
END_REGION

REGION Network 6: Debloquer consigne
   RUNG wire#powerrail
      Contact( "Bits_Globaux".x_En_service )
      Coil( #DB_Variateur.Cmd.DebloqConsigne )
   END_RUNG
   // the same network as SCL:
   #DB_Variateur.Cmd.DebloqConsigne := "Bits_Globaux".x_En_service;
END_REGION

REGION Network 7: Inversion de sens
   RUNG wire#powerrail
      Contact( #InversionSens )
      Coil( #DB_Variateur.Cmd.InversionConsigne )
   END_RUNG
   // the same network as SCL:
   #DB_Variateur.Cmd.InversionConsigne := #InversionSens;
END_REGION

REGION Network 8: Consigne manu
   RUNG wire#powerrail
      Contact( "Bits_Globaux".x_En_manu )
      { S7_Templates := "[SrcType := Int, DestType := Real]" } Normalize(min := int#0, value := #"Vitesse MANU", max := int#1380, out => #ResultNorm_sp)
      { S7_Templates := "[SrcType := Real, DestType := Int]" } Scale(min := 0, value := #ResultNorm_sp, max := 16384, out => #ResultScale_sp)
      Move(in := #ResultScale_sp, out1 => #DB_Variateur.Cmd.Consigne)
   END_RUNG
   // the same network as SCL:
   IF "Bits_Globaux".x_En_manu THEN
       #ResultNorm_sp := NORM_X(MIN := int#0, VALUE := #"Vitesse MANU", MAX := int#1380);
       #ResultScale_sp := SCALE_X(MIN := 0, VALUE := #ResultNorm_sp, MAX := 16384);
       #DB_Variateur.Cmd.Consigne := #ResultScale_sp;
   END_IF;
END_REGION

REGION Network 9: Consigne auto
   RUNG wire#powerrail
      Contact( "I_En_Automatique" )
      { S7_Templates := "[SrcType := Int, DestType := Real]" } Normalize(min := int#0, value := #"Vitesse AUTO", max := int#1380, out => #ResultNorm_sp)
      { S7_Templates := "[SrcType := Real, DestType := Int]" } Scale(min := 0, value := #ResultNorm_sp, max := 16384, out => #ResultScale_sp)
      Move(in := #ResultScale_sp, out1 => #DB_Variateur.Cmd.Consigne)
   END_RUNG
   // the same network as SCL:
   IF "I_En_Automatique" THEN
       #ResultNorm_sp := NORM_X(MIN := int#0, VALUE := #"Vitesse AUTO", MAX := int#1380);
       #ResultScale_sp := SCALE_X(MIN := 0, VALUE := #ResultNorm_sp, MAX := 16384);
       #DB_Variateur.Cmd.Consigne := #ResultScale_sp;
   END_IF;
END_REGION

REGION Network 10: Acquiter defauts
   RUNG wire#powerrail
      Contact( #Ack_defaut )
      wire#w1
      Coil( #DB_Variateur.Cmd.AcquitDefaut )
   END_RUNG
   RUNG wire#powerrail
      Contact( #Rearmement )
   END_RUNG wire#w1
   // the same network as SCL:
   #DB_Variateur.Cmd.AcquitDefaut := #Ack_defaut OR #Rearmement;
END_REGION

REGION Network 11: Marche moteur
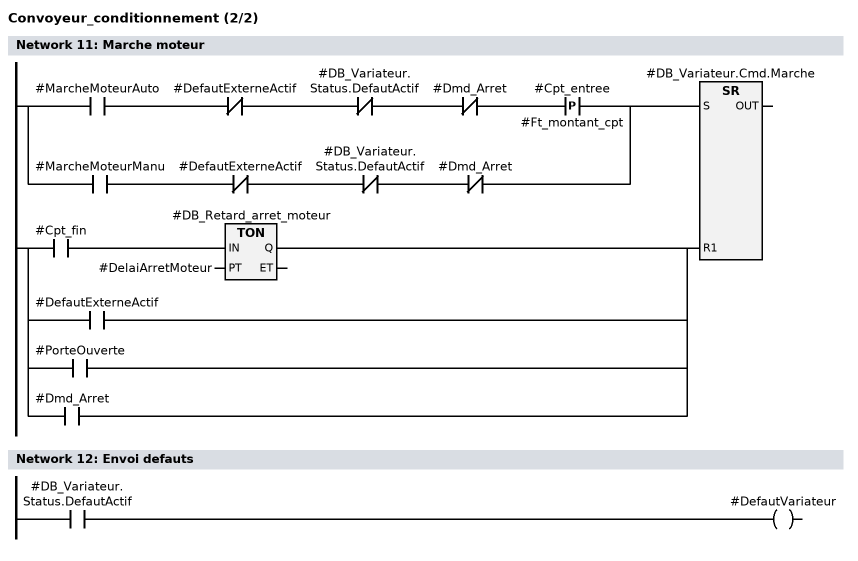
   #_w1 := #MarcheMoteurAuto AND NOT #DefautExterneActif AND NOT #DB_Variateur.Status.DefautActif AND NOT #Dmd_Arret AND #Cpt_entree AND NOT #Ft_montant_cpt;   // rising edge of #Cpt_entree
   #Ft_montant_cpt := #Cpt_entree;
   #DB_Retard_arret_moteur(IN := #Cpt_fin, PT := #DelaiArretMoteur);   // TON
   IF #_w1 OR (#MarcheMoteurManu AND NOT #DefautExterneActif AND NOT #DB_Variateur.Status.DefautActif AND NOT #Dmd_Arret) THEN
       #DB_Variateur.Cmd.Marche := TRUE;   // SR flip-flop
   END_IF;
   IF #DB_Retard_arret_moteur.Q OR #DefautExterneActif OR #PorteOuverte OR #Dmd_Arret THEN
       #DB_Variateur.Cmd.Marche := FALSE;
   END_IF;
END_REGION

REGION Network 12: Envoi defauts
   RUNG wire#powerrail
      Contact( #DB_Variateur.Status.DefautActif )
      Coil( #DefautVariateur )
   END_RUNG
   // the same network as SCL:
   #DefautVariateur := #DB_Variateur.Status.DefautActif;
END_REGION
END_FUNCTION_BLOCK

FUNCTION_BLOCK "Gestion_Convoyeurs"   // FB7, LAD
TITLE = Gestion des convoyeurs
{ S7_Optimized_Access := 'TRUE' }
VERSION : 0.1
   VAR
      Convoyeur_1 : "Convoyeur_conditionnement";
      Convoyeur_2 : "Convoyeur_conditionnement";
      Convoyeur_3 : "Convoyeur_conditionnement";
   END_VAR
BEGIN

REGION Network 1: Commande convoyeur 1
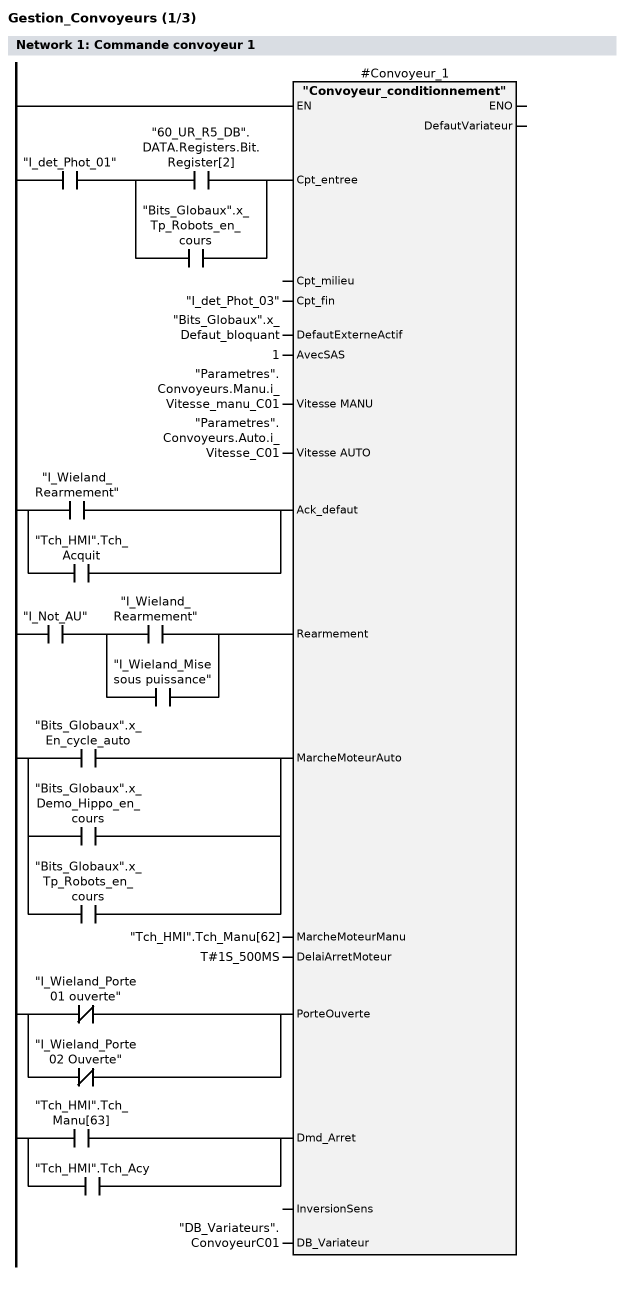
   RUNG wire#powerrail
      #Convoyeur_1(Cpt_entree := wire#w2, Ack_defaut := wire#w3, Rearmement := wire#w5, MarcheMoteurAuto := wire#w6, PorteOuverte := wire#w7, Dmd_Arret := wire#w8, Cpt_milieu :=, Cpt_fin := "I_det_Phot_03", DefautExterneActif := "Bits_Globaux".x_Defaut_bloquant, AvecSAS := 1, "Vitesse MANU" := "Parametres".Convoyeurs.Manu.i_Vitesse_manu_C01, "Vitesse AUTO" := "Parametres".Convoyeurs.Auto.i_Vitesse_C01, MarcheMoteurManu := "Tch_HMI".Tch_Manu[62], DelaiArretMoteur := T#1S_500MS, InversionSens :=, DB_Variateur := "DB_Variateurs".ConvoyeurC01, DefautVariateur =>)
   END_RUNG
   RUNG wire#powerrail
      Contact( "I_det_Phot_01" )
      wire#w1
      Contact( "60_UR_R5_DB".DATA.Registers.Bit.Register[2] )
   END_RUNG wire#w2
   RUNG wire#w1
      Contact( "Bits_Globaux".x_Tp_Robots_en_cours )
   END_RUNG wire#w2
   RUNG wire#powerrail
      Contact( "I_Wieland_Rearmement" )
   END_RUNG wire#w3
   RUNG wire#powerrail
      Contact( "Tch_HMI".Tch_Acquit )
   END_RUNG wire#w3
   RUNG wire#powerrail
      Contact( "I_Not_AU" )
      wire#w4
      Contact( "I_Wieland_Rearmement" )
   END_RUNG wire#w5
   RUNG wire#w4
      Contact( "I_Wieland_Mise sous puissance" )
   END_RUNG wire#w5
   RUNG wire#powerrail
      Contact( "Bits_Globaux".x_En_cycle_auto )
   END_RUNG wire#w6
   RUNG wire#powerrail
      Contact( "Bits_Globaux".x_Demo_Hippo_en_cours )
   END_RUNG wire#w6
   RUNG wire#powerrail
      Contact( "Bits_Globaux".x_Tp_Robots_en_cours )
   END_RUNG wire#w6
   RUNG wire#powerrail
      I_Contact( "I_Wieland_Porte 01 ouverte" )
   END_RUNG wire#w7
   RUNG wire#powerrail
      I_Contact( "I_Wieland_Porte 02 Ouverte" )
   END_RUNG wire#w7
   RUNG wire#powerrail
      Contact( "Tch_HMI".Tch_Manu[63] )
   END_RUNG wire#w8
   RUNG wire#powerrail
      Contact( "Tch_HMI".Tch_Acy )
   END_RUNG wire#w8
   // the same network as SCL:
   #Convoyeur_1(Cpt_entree := "I_det_Phot_01" AND ("60_UR_R5_DB".DATA.Registers.Bit.Register[2] OR "Bits_Globaux".x_Tp_Robots_en_cours),   // "Convoyeur_conditionnement"
                Cpt_fin := "I_det_Phot_03",
                DefautExterneActif := "Bits_Globaux".x_Defaut_bloquant,
                AvecSAS := 1,
                "Vitesse MANU" := "Parametres".Convoyeurs.Manu.i_Vitesse_manu_C01,
                "Vitesse AUTO" := "Parametres".Convoyeurs.Auto.i_Vitesse_C01,
                Ack_defaut := "I_Wieland_Rearmement" OR "Tch_HMI".Tch_Acquit,
                Rearmement := "I_Not_AU" AND ("I_Wieland_Rearmement" OR "I_Wieland_Mise sous puissance"),
                MarcheMoteurAuto := "Bits_Globaux".x_En_cycle_auto OR "Bits_Globaux".x_Demo_Hippo_en_cours OR "Bits_Globaux".x_Tp_Robots_en_cours,
                MarcheMoteurManu := "Tch_HMI".Tch_Manu[62],
                DelaiArretMoteur := T#1S_500MS,
                PorteOuverte := NOT "I_Wieland_Porte 01 ouverte" OR NOT "I_Wieland_Porte 02 Ouverte",
                Dmd_Arret := "Tch_HMI".Tch_Manu[63] OR "Tch_HMI".Tch_Acy,
                DB_Variateur := "DB_Variateurs".ConvoyeurC01);
END_REGION

REGION Network 2: Commande convoyeur 2
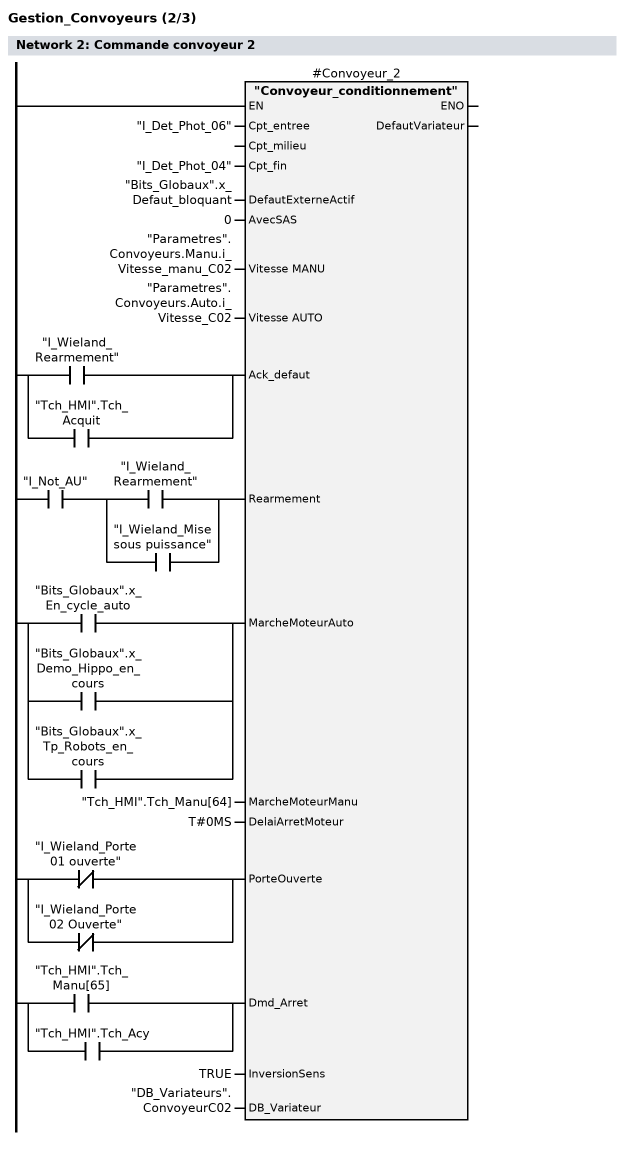
   RUNG wire#powerrail
      #Convoyeur_2(Ack_defaut := wire#w1, Rearmement := wire#w3, MarcheMoteurAuto := wire#w4, PorteOuverte := wire#w5, Dmd_Arret := wire#w6, Cpt_entree := "I_Det_Phot_06", Cpt_milieu :=, Cpt_fin := "I_Det_Phot_04", DefautExterneActif := "Bits_Globaux".x_Defaut_bloquant, AvecSAS := 0, "Vitesse MANU" := "Parametres".Convoyeurs.Manu.i_Vitesse_manu_C02, "Vitesse AUTO" := "Parametres".Convoyeurs.Auto.i_Vitesse_C02, MarcheMoteurManu := "Tch_HMI".Tch_Manu[64], DelaiArretMoteur := T#0MS, InversionSens := TRUE, DB_Variateur := "DB_Variateurs".ConvoyeurC02, DefautVariateur =>)
   END_RUNG
   RUNG wire#powerrail
      Contact( "I_Wieland_Rearmement" )
   END_RUNG wire#w1
   RUNG wire#powerrail
      Contact( "Tch_HMI".Tch_Acquit )
   END_RUNG wire#w1
   RUNG wire#powerrail
      Contact( "I_Not_AU" )
      wire#w2
      Contact( "I_Wieland_Rearmement" )
   END_RUNG wire#w3
   RUNG wire#w2
      Contact( "I_Wieland_Mise sous puissance" )
   END_RUNG wire#w3
   RUNG wire#powerrail
      Contact( "Bits_Globaux".x_En_cycle_auto )
   END_RUNG wire#w4
   RUNG wire#powerrail
      Contact( "Bits_Globaux".x_Demo_Hippo_en_cours )
   END_RUNG wire#w4
   RUNG wire#powerrail
      Contact( "Bits_Globaux".x_Tp_Robots_en_cours )
   END_RUNG wire#w4
   RUNG wire#powerrail
      I_Contact( "I_Wieland_Porte 01 ouverte" )
   END_RUNG wire#w5
   RUNG wire#powerrail
      I_Contact( "I_Wieland_Porte 02 Ouverte" )
   END_RUNG wire#w5
   RUNG wire#powerrail
      Contact( "Tch_HMI".Tch_Manu[65] )
   END_RUNG wire#w6
   RUNG wire#powerrail
      Contact( "Tch_HMI".Tch_Acy )
   END_RUNG wire#w6
   // the same network as SCL:
   #Convoyeur_2(Cpt_entree := "I_Det_Phot_06",   // "Convoyeur_conditionnement"
                Cpt_fin := "I_Det_Phot_04",
                DefautExterneActif := "Bits_Globaux".x_Defaut_bloquant,
                AvecSAS := 0,
                "Vitesse MANU" := "Parametres".Convoyeurs.Manu.i_Vitesse_manu_C02,
                "Vitesse AUTO" := "Parametres".Convoyeurs.Auto.i_Vitesse_C02,
                Ack_defaut := "I_Wieland_Rearmement" OR "Tch_HMI".Tch_Acquit,
                Rearmement := "I_Not_AU" AND ("I_Wieland_Rearmement" OR "I_Wieland_Mise sous puissance"),
                MarcheMoteurAuto := "Bits_Globaux".x_En_cycle_auto OR "Bits_Globaux".x_Demo_Hippo_en_cours OR "Bits_Globaux".x_Tp_Robots_en_cours,
                MarcheMoteurManu := "Tch_HMI".Tch_Manu[64],
                DelaiArretMoteur := T#0MS,
                PorteOuverte := NOT "I_Wieland_Porte 01 ouverte" OR NOT "I_Wieland_Porte 02 Ouverte",
                Dmd_Arret := "Tch_HMI".Tch_Manu[65] OR "Tch_HMI".Tch_Acy,
                InversionSens := TRUE,
                DB_Variateur := "DB_Variateurs".ConvoyeurC02);
END_REGION

REGION Network 3: Commande convoyeur 3
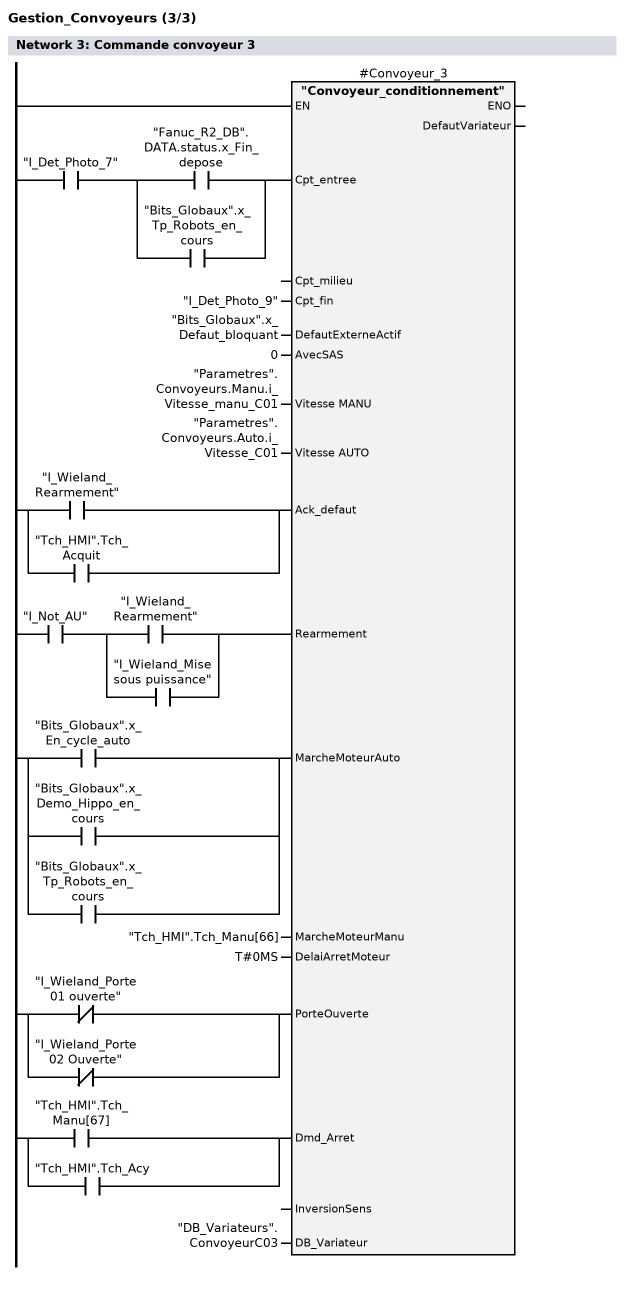
   RUNG wire#powerrail
      #Convoyeur_3(Cpt_entree := wire#w2, Ack_defaut := wire#w3, Rearmement := wire#w5, MarcheMoteurAuto := wire#w6, PorteOuverte := wire#w7, Dmd_Arret := wire#w8, Cpt_milieu :=, Cpt_fin := "I_Det_Photo_9", DefautExterneActif := "Bits_Globaux".x_Defaut_bloquant, AvecSAS := 0, "Vitesse MANU" := "Parametres".Convoyeurs.Manu.i_Vitesse_manu_C01, "Vitesse AUTO" := "Parametres".Convoyeurs.Auto.i_Vitesse_C01, MarcheMoteurManu := "Tch_HMI".Tch_Manu[66], DelaiArretMoteur := T#0MS, InversionSens :=, DB_Variateur := "DB_Variateurs".ConvoyeurC03, DefautVariateur =>)
   END_RUNG
   RUNG wire#powerrail
      Contact( "I_Det_Photo_7" )
      wire#w1
      Contact( "Fanuc_R2_DB".DATA.status.x_Fin_depose )
   END_RUNG wire#w2
   RUNG wire#w1
      Contact( "Bits_Globaux".x_Tp_Robots_en_cours )
   END_RUNG wire#w2
   RUNG wire#powerrail
      Contact( "I_Wieland_Rearmement" )
   END_RUNG wire#w3
   RUNG wire#powerrail
      Contact( "Tch_HMI".Tch_Acquit )
   END_RUNG wire#w3
   RUNG wire#powerrail
      Contact( "I_Not_AU" )
      wire#w4
      Contact( "I_Wieland_Rearmement" )
   END_RUNG wire#w5
   RUNG wire#w4
      Contact( "I_Wieland_Mise sous puissance" )
   END_RUNG wire#w5
   RUNG wire#powerrail
      Contact( "Bits_Globaux".x_En_cycle_auto )
   END_RUNG wire#w6
   RUNG wire#powerrail
      Contact( "Bits_Globaux".x_Demo_Hippo_en_cours )
   END_RUNG wire#w6
   RUNG wire#powerrail
      Contact( "Bits_Globaux".x_Tp_Robots_en_cours )
   END_RUNG wire#w6
   RUNG wire#powerrail
      I_Contact( "I_Wieland_Porte 01 ouverte" )
   END_RUNG wire#w7
   RUNG wire#powerrail
      I_Contact( "I_Wieland_Porte 02 Ouverte" )
   END_RUNG wire#w7
   RUNG wire#powerrail
      Contact( "Tch_HMI".Tch_Manu[67] )
   END_RUNG wire#w8
   RUNG wire#powerrail
      Contact( "Tch_HMI".Tch_Acy )
   END_RUNG wire#w8
   // the same network as SCL:
   #Convoyeur_3(Cpt_entree := "I_Det_Photo_7" AND ("Fanuc_R2_DB".DATA.status.x_Fin_depose OR "Bits_Globaux".x_Tp_Robots_en_cours),   // "Convoyeur_conditionnement"
                Cpt_fin := "I_Det_Photo_9",
                DefautExterneActif := "Bits_Globaux".x_Defaut_bloquant,
                AvecSAS := 0,
                "Vitesse MANU" := "Parametres".Convoyeurs.Manu.i_Vitesse_manu_C01,
                "Vitesse AUTO" := "Parametres".Convoyeurs.Auto.i_Vitesse_C01,
                Ack_defaut := "I_Wieland_Rearmement" OR "Tch_HMI".Tch_Acquit,
                Rearmement := "I_Not_AU" AND ("I_Wieland_Rearmement" OR "I_Wieland_Mise sous puissance"),
                MarcheMoteurAuto := "Bits_Globaux".x_En_cycle_auto OR "Bits_Globaux".x_Demo_Hippo_en_cours OR "Bits_Globaux".x_Tp_Robots_en_cours,
                MarcheMoteurManu := "Tch_HMI".Tch_Manu[66],
                DelaiArretMoteur := T#0MS,
                PorteOuverte := NOT "I_Wieland_Porte 01 ouverte" OR NOT "I_Wieland_Porte 02 Ouverte",
                Dmd_Arret := "Tch_HMI".Tch_Manu[67] OR "Tch_HMI".Tch_Acy,
                DB_Variateur := "DB_Variateurs".ConvoyeurC03);
END_REGION
END_FUNCTION_BLOCK

// folder: 5-Cellule_conditionnement/Fanuc_R1

FUNCTION_BLOCK "Fanuc_R1"   // FB3, LAD
{ S7_Optimized_Access := 'TRUE' }
VERSION : 0.1
   VAR
      DATA : "Fanuc_Robot";
      Front_montant_Init : Bool;
   END_VAR
BEGIN

REGION Network 1: Grafcet
END_REGION

REGION Network 2: Gestion defauts
END_REGION

REGION Network 3: Post traitement
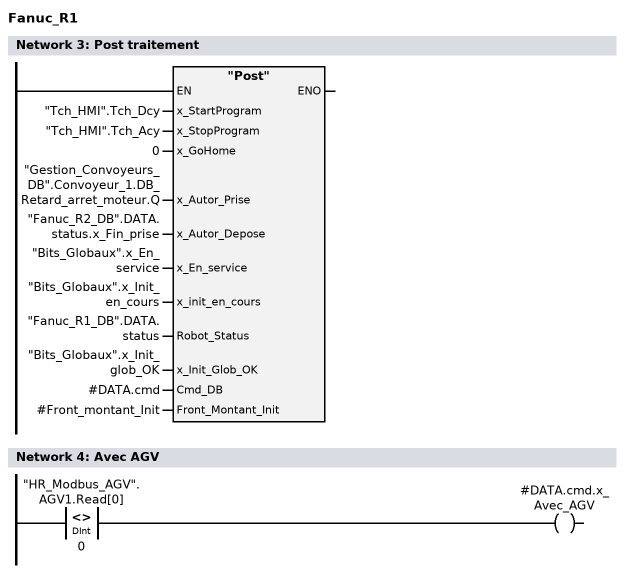
   RUNG wire#powerrail
      "Post"(x_StartProgram := "Tch_HMI".Tch_Dcy, x_StopProgram := "Tch_HMI".Tch_Acy, x_GoHome := 0, x_Autor_Prise := "Gestion_Convoyeurs_DB".Convoyeur_1.DB_Retard_arret_moteur.Q, x_Autor_Depose := "Fanuc_R2_DB".DATA.status.x_Fin_prise, x_En_service := "Bits_Globaux".x_En_service, x_init_en_cours := "Bits_Globaux".x_Init_en_cours, Robot_Status := "Fanuc_R1_DB".DATA.status, x_Init_Glob_OK := "Bits_Globaux".x_Init_glob_OK, Cmd_DB := #DATA.cmd, Front_Montant_Init := #Front_montant_Init)
   END_RUNG
   // the same network as SCL:
   "Post"(x_StartProgram := "Tch_HMI".Tch_Dcy,
          x_StopProgram := "Tch_HMI".Tch_Acy,
          x_GoHome := 0,
          x_Autor_Prise := "Gestion_Convoyeurs_DB".Convoyeur_1.DB_Retard_arret_moteur.Q,
          x_Autor_Depose := "Fanuc_R2_DB".DATA.status.x_Fin_prise,
          x_En_service := "Bits_Globaux".x_En_service,
          x_init_en_cours := "Bits_Globaux".x_Init_en_cours,
          Robot_Status := "Fanuc_R1_DB".DATA.status,
          x_Init_Glob_OK := "Bits_Globaux".x_Init_glob_OK,
          Cmd_DB := #DATA.cmd,
          Front_Montant_Init := #Front_montant_Init);
END_REGION

REGION Network 4: Avec AGV
   RUNG wire#powerrail
      { S7_Templates := "SrcType := DInt" } NE_Contact(in1 := "HR_Modbus_AGV".AGV1.Read[0], in2 := 0)
      Coil( #DATA.cmd.x_Avec_AGV )
   END_RUNG
   // the same network as SCL:
   #DATA.cmd.x_Avec_AGV := "HR_Modbus_AGV".AGV1.Read[0] <> 0;
END_REGION
END_FUNCTION_BLOCK

FUNCTION "Post" : Void   // FC9, LAD
TITLE = POST Fanuc
{ S7_Optimized_Access := 'TRUE' }
VERSION : 0.1
   VAR_INPUT
      x_StartProgram : Bool;
      x_StopProgram : Bool;
      x_GoHome : Bool;
      x_Autor_Prise : Bool;
      x_Autor_Depose : Bool;
      x_En_service : Bool;
      x_init_en_cours : Bool;
      Robot_Status : "Fanuc_status";
      x_Init_Glob_OK : Bool;
   END_VAR
   VAR_IN_OUT
      Cmd_DB : "Fanuc_cmd";
      Front_Montant_Init : Bool;
   END_VAR
BEGIN

REGION Network 1: IMSTP
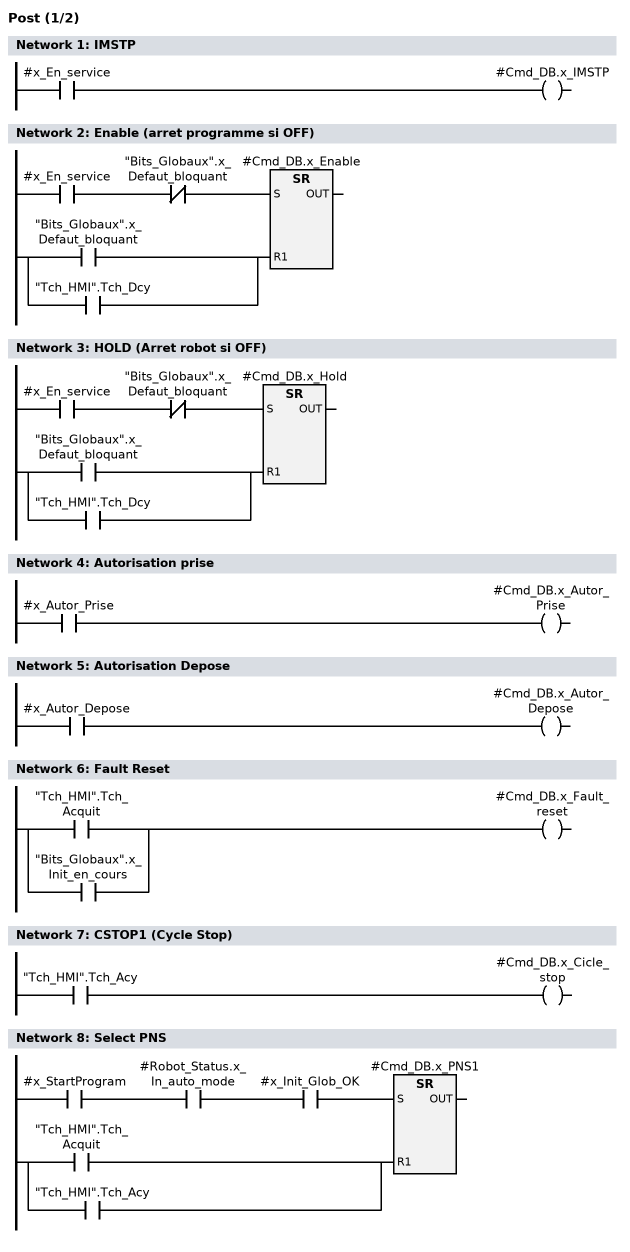
   RUNG wire#powerrail
      Contact( #x_En_service )
      Coil( #Cmd_DB.x_IMSTP )
   END_RUNG
   // the same network as SCL:
   #Cmd_DB.x_IMSTP := #x_En_service;
END_REGION

REGION Network 2: Enable (arret programme si OFF)
   RUNG wire#powerrail
      Contact( #x_En_service )
      I_Contact( "Bits_Globaux".x_Defaut_bloquant )
      S_SR(operand := #Cmd_DB.x_Enable, r1 := wire#w1)
   END_RUNG
   RUNG wire#powerrail
      Contact( "Bits_Globaux".x_Defaut_bloquant )
   END_RUNG wire#w1
   RUNG wire#powerrail
      Contact( "Tch_HMI".Tch_Dcy )
   END_RUNG wire#w1
   // the same network as SCL:
   IF #x_En_service AND NOT "Bits_Globaux".x_Defaut_bloquant THEN
       #Cmd_DB.x_Enable := TRUE;   // SR flip-flop
   END_IF;
   IF "Bits_Globaux".x_Defaut_bloquant OR "Tch_HMI".Tch_Dcy THEN #Cmd_DB.x_Enable := FALSE; END_IF;
END_REGION

REGION Network 3: HOLD (Arret robot si OFF)
   RUNG wire#powerrail
      Contact( #x_En_service )
      I_Contact( "Bits_Globaux".x_Defaut_bloquant )
      S_SR(operand := #Cmd_DB.x_Hold, r1 := wire#w1)
   END_RUNG
   RUNG wire#powerrail
      Contact( "Bits_Globaux".x_Defaut_bloquant )
   END_RUNG wire#w1
   RUNG wire#powerrail
      Contact( "Tch_HMI".Tch_Dcy )
   END_RUNG wire#w1
   // the same network as SCL:
   IF #x_En_service AND NOT "Bits_Globaux".x_Defaut_bloquant THEN
       #Cmd_DB.x_Hold := TRUE;   // SR flip-flop
   END_IF;
   IF "Bits_Globaux".x_Defaut_bloquant OR "Tch_HMI".Tch_Dcy THEN #Cmd_DB.x_Hold := FALSE; END_IF;
END_REGION

REGION Network 4: Autorisation prise
   RUNG wire#powerrail
      Contact( #x_Autor_Prise )
      Coil( #Cmd_DB.x_Autor_Prise )
   END_RUNG
   // the same network as SCL:
   #Cmd_DB.x_Autor_Prise := #x_Autor_Prise;
END_REGION

REGION Network 5: Autorisation Depose
   RUNG wire#powerrail
      Contact( #x_Autor_Depose )
      Coil( #Cmd_DB.x_Autor_Depose )
   END_RUNG
   // the same network as SCL:
   #Cmd_DB.x_Autor_Depose := #x_Autor_Depose;
END_REGION

REGION Network 6: Fault Reset
   RUNG wire#powerrail
      Contact( "Tch_HMI".Tch_Acquit )
      wire#w1
      Coil( #Cmd_DB.x_Fault_reset )
   END_RUNG
   RUNG wire#powerrail
      Contact( "Bits_Globaux".x_Init_en_cours )
   END_RUNG wire#w1
   // the same network as SCL:
   #Cmd_DB.x_Fault_reset := "Tch_HMI".Tch_Acquit OR "Bits_Globaux".x_Init_en_cours;
END_REGION

REGION Network 7: CSTOP1 (Cycle Stop)
   RUNG wire#powerrail
      Contact( "Tch_HMI".Tch_Acy )
      Coil( #Cmd_DB.x_Cicle_stop )
   END_RUNG
   // the same network as SCL:
   #Cmd_DB.x_Cicle_stop := "Tch_HMI".Tch_Acy;
END_REGION

REGION Network 8: Select PNS
   RUNG wire#powerrail
      Contact( #x_StartProgram )
      Contact( #Robot_Status.x_In_auto_mode )
      Contact( #x_Init_Glob_OK )
      S_SR(operand := #Cmd_DB.x_PNS1, r1 := wire#w1)
   END_RUNG
   RUNG wire#powerrail
      Contact( "Tch_HMI".Tch_Acquit )
   END_RUNG wire#w1
   RUNG wire#powerrail
      Contact( "Tch_HMI".Tch_Acy )
   END_RUNG wire#w1
   // the same network as SCL:
   IF #x_StartProgram AND #Robot_Status.x_In_auto_mode AND #x_Init_Glob_OK THEN
       #Cmd_DB.x_PNS1 := TRUE;   // SR flip-flop
   END_IF;
   IF "Tch_HMI".Tch_Acquit OR "Tch_HMI".Tch_Acy THEN #Cmd_DB.x_PNS1 := FALSE; END_IF;
END_REGION

REGION Network 9: Start PNS program
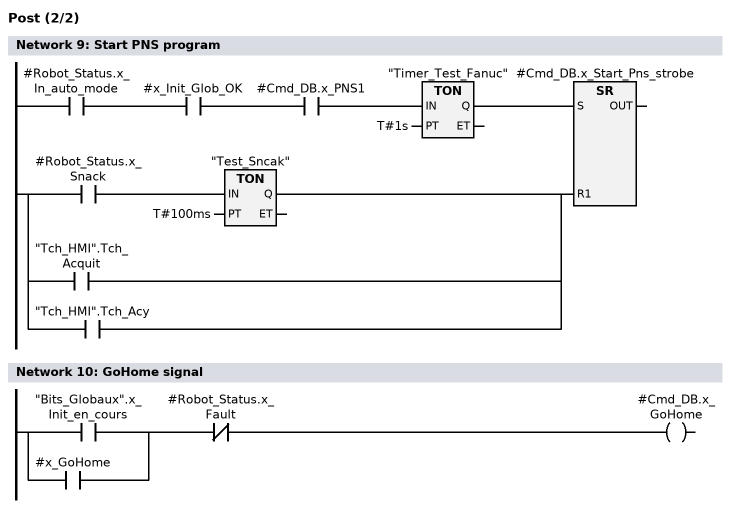
   "Timer_Test_Fanuc".TON(IN := #Robot_Status.x_In_auto_mode AND #x_Init_Glob_OK AND #Cmd_DB.x_PNS1, PT := T#1s);
   "Test_Sncak".TON(IN := #Robot_Status.x_Snack, PT := T#100ms);
   IF "Timer_Test_Fanuc".Q THEN
       #Cmd_DB.x_Start_Pns_strobe := TRUE;   // SR flip-flop
   END_IF;
   IF "Test_Sncak".Q OR "Tch_HMI".Tch_Acquit OR "Tch_HMI".Tch_Acy THEN
       #Cmd_DB.x_Start_Pns_strobe := FALSE;
   END_IF;
END_REGION

REGION Network 10: GoHome signal
   RUNG wire#powerrail
      Contact( "Bits_Globaux".x_Init_en_cours )
      wire#w1
      I_Contact( #Robot_Status.x_Fault )
      Coil( #Cmd_DB.x_GoHome )
   END_RUNG
   RUNG wire#powerrail
      Contact( #x_GoHome )
   END_RUNG wire#w1
   // the same network as SCL:
   #Cmd_DB.x_GoHome := ("Bits_Globaux".x_Init_en_cours OR #x_GoHome) AND NOT #Robot_Status.x_Fault;
END_REGION
END_FUNCTION

// folder: 5-Cellule_conditionnement/Fanuc_R2

FUNCTION_BLOCK "Fanuc_R2"   // FB5, LAD
{ S7_Optimized_Access := 'TRUE' }
VERSION : 0.1
   VAR
      DATA : "Fanuc_Robot";
      Front_Montant_Init : Bool;
   END_VAR
BEGIN

REGION Network 2: POST Traitement FANUC R2
